   // ---------- 网络 20 ----------
   // 标题：*************故障计数（包含水平钻超时，凿超时，低电流，打孔深度超限）***********************
   // 注释：VisualChiseling No Sloping Hammer, added not  DB2500.DBX30.0  and #DrillHorizontal.StopDrill_Ack (in Network End) by WXY, 20220726
   // 含义：调用计数器实例 "Timer_DrilEndPos".TON（上升沿计数，当前值写入 CV）
   "Timer_DrilEndPos".TON(IN := (((((#HorDrillStep.S20 AND NOT (#HorDrillStep.S22)) OR ((#HorDrillStep.S22 AND NOT (#HorDrillStep.S25)) AND NOT ("DB2500 Visual Chiseling".VisualChiselingMode))) AND "DB1900_Communication_PC".Para.ProduceMode3) AND "DB720_KuKa_MainCtrl".StatusIn.do_DrilEnd_Pos) AND ("DB1900_Communication_PC".Recv.Current_2 < "DB1900_Communication_PC".Para.CurrentMinLimit)),
                          PT := T#2s);
   // 含义：条件 "Timer_DrilEndPos".Q 成立时，将 TRUE 传送到 "DB2500 Visual Chiseling".VChiselEndPos
   IF "Timer_DrilEndPos".Q THEN
       "DB2500 Visual Chiseling".VChiselEndPos := TRUE;
   END_IF;
   // 含义：条件 "Timer_DrilEndPos".Q 成立时，将 ("DB1042_Timer".HCLowTimeOutTimes + 1) 传送到 "DB1042_Timer".HCLowTimeOutTimes
   IF "Timer_DrilEndPos".Q THEN
       "DB1042_Timer".HCLowTimeOutTimes := ("DB1042_Timer".HCLowTimeOutTimes + 1);
   END_IF;
   // 含义：条件 ((((((#HorDrillStep.S20 AND NOT (#HorDrillStep.S22)) OR ((#HorDrillStep.S22 AND NOT (#HorDrillStep.S25)) AND NOT ("DB2500 Visual Chiseling".VisualChiselingMode))) AND "DB1900_Communication_PC".Para.ProduceMode3) AND ("DB1900_Communication_PC".Recv.Current_2 > "DB1900_Communication_PC".Para.CurrentMinLimit))) AND ("DB1900_Communication_PC".Recv.Current_2 < "DB1900_Communication_PC".Para.CurrentMaxLimit)) 成立时，将 0 传送到 "DB1042_Timer".HCLowTimeOutTimes
   IF ((((((#HorDrillStep.S20 AND NOT (#HorDrillStep.S22)) OR ((#HorDrillStep.S22 AND NOT (#HorDrillStep.S25)) AND NOT ("DB2500 Visual Chiseling".VisualChiselingMode))) AND "DB1900_Communication_PC".Para.ProduceMode3) AND ("DB1900_Communication_PC".Recv.Current_2 > "DB1900_Communication_PC".Para.CurrentMinLimit))) AND ("DB1900_Communication_PC".Recv.Current_2 < "DB1900_Communication_PC".Para.CurrentMaxLimit)) THEN
       "DB1042_Timer".HCLowTimeOutTimes := 0;
   END_IF;
   // 含义：条件 (((((#HorDrillStep.S20 AND NOT (#HorDrillStep.S22)) OR ((#HorDrillStep.S22 AND NOT (#HorDrillStep.S25)) AND NOT ("DB2500 Visual Chiseling".VisualChiselingMode))) AND "DB1900_Communication_PC".Para.ProduceMode3) AND "DB1042_Timer".HDrillEndTime.Q) OR ((((#HorDrillStep.S20 AND NOT (#HorDrillStep.S22)) OR ((#HorDrillStep.S22 AND NOT (#HorDrillStep.S25)) AND NOT ("DB2500 Visual Chiseling".VisualChiselingMode))) AND "DB1900_Communication_PC".Para.ProduceMode3) AND "DB1042_Timer".GougeTimeOut.Q) OR ((((#HorDrillStep.S20 AND NOT (#HorDrillStep.S22)) OR ((#HorDrillStep.S22 AND NOT (#HorDrillStep.S25)) AND NOT ("DB2500 Visual Chiseling".VisualChiselingMode))) AND "DB1900_Communication_PC".Para.ProduceMode3) AND "DB1042_Timer".CurrentLowTimeOut.Q) OR ((((#HorDrillStep.S20 AND NOT (#HorDrillStep.S22)) OR ((#HorDrillStep.S22 AND NOT (#HorDrillStep.S25)) AND NOT ("DB2500 Visual Chiseling".VisualChiselingMode))) AND "DB1900_Communication_PC".Para.ProduceMode3) AND "DB1042_Timer".CurrentHighTimeOut.Q) OR (((((#HorDrillStep.S20 AND NOT (#HorDrillStep.S22)) OR ((#HorDrillStep.S22 AND NOT (#HorDrillStep.S25)) AND NOT ("DB2500 Visual Chiseling".VisualChiselingMode))) AND "DB1900_Communication_PC".Para.ProduceMode3) AND ("DB1900_Communication_PC".Send.ScrLen >= "DB1900_Communication_PC".Para.DrillDepth))) OR ((((#HorDrillStep.S20 AND NOT (#HorDrillStep.S22)) OR ((#HorDrillStep.S22 AND NOT (#HorDrillStep.S25)) AND NOT ("DB2500 Visual Chiseling".VisualChiselingMode))) AND "DB1900_Communication_PC".Para.ProduceMode3) AND "DB2500 Visual Chiseling".VChiselEndPos)) AND NOT ("DB720_KuKa_MainCtrl".StatusIn.do_ChiselCylinderExt) 成立时，将 0.1 传送到 "DB1080_Component".Aux.Pressure
   IF (((((#HorDrillStep.S20 AND NOT (#HorDrillStep.S22)) OR ((#HorDrillStep.S22 AND NOT (#HorDrillStep.S25)) AND NOT ("DB2500 Visual Chiseling".VisualChiselingMode))) AND "DB1900_Communication_PC".Para.ProduceMode3) AND "DB1042_Timer".HDrillEndTime.Q) OR ((((#HorDrillStep.S20 AND NOT (#HorDrillStep.S22)) OR ((#HorDrillStep.S22 AND NOT (#HorDrillStep.S25)) AND NOT ("DB2500 Visual Chiseling".VisualChiselingMode))) AND "DB1900_Communication_PC".Para.ProduceMode3) AND "DB1042_Timer".GougeTimeOut.Q) OR ((((#HorDrillStep.S20 AND NOT (#HorDrillStep.S22)) OR ((#HorDrillStep.S22 AND NOT (#HorDrillStep.S25)) AND NOT ("DB2500 Visual Chiseling".VisualChiselingMode))) AND "DB1900_Communication_PC".Para.ProduceMode3) AND "DB1042_Timer".CurrentLowTimeOut.Q) OR ((((#HorDrillStep.S20 AND NOT (#HorDrillStep.S22)) OR ((#HorDrillStep.S22 AND NOT (#HorDrillStep.S25)) AND NOT ("DB2500 Visual Chiseling".VisualChiselingMode))) AND "DB1900_Communication_PC".Para.ProduceMode3) AND "DB1042_Timer".CurrentHighTimeOut.Q) OR (((((#HorDrillStep.S20 AND NOT (#HorDrillStep.S22)) OR ((#HorDrillStep.S22 AND NOT (#HorDrillStep.S25)) AND NOT ("DB2500 Visual Chiseling".VisualChiselingMode))) AND "DB1900_Communication_PC".Para.ProduceMode3) AND ("DB1900_Communication_PC".Send.ScrLen >= "DB1900_Communication_PC".Para.DrillDepth))) OR ((((#HorDrillStep.S20 AND NOT (#HorDrillStep.S22)) OR ((#HorDrillStep.S22 AND NOT (#HorDrillStep.S25)) AND NOT ("DB2500 Visual Chiseling".VisualChiselingMode))) AND "DB1900_Communication_PC".Para.ProduceMode3) AND "DB2500 Visual Chiseling".VChiselEndPos)) AND NOT ("DB720_KuKa_MainCtrl".StatusIn.do_ChiselCylinderExt) THEN
       "DB1080_Component".Aux.Pressure := 0.1;
   END_IF;
   // 含义：条件 (((((#HorDrillStep.S20 AND NOT (#HorDrillStep.S22)) OR ((#HorDrillStep.S22 AND NOT (#HorDrillStep.S25)) AND NOT ("DB2500 Visual Chiseling".VisualChiselingMode))) AND "DB1900_Communication_PC".Para.ProduceMode3) AND "DB1042_Timer".HDrillEndTime.Q) OR ((((#HorDrillStep.S20 AND NOT (#HorDrillStep.S22)) OR ((#HorDrillStep.S22 AND NOT (#HorDrillStep.S25)) AND NOT ("DB2500 Visual Chiseling".VisualChiselingMode))) AND "DB1900_Communication_PC".Para.ProduceMode3) AND "DB1042_Timer".GougeTimeOut.Q) OR ((((#HorDrillStep.S20 AND NOT (#HorDrillStep.S22)) OR ((#HorDrillStep.S22 AND NOT (#HorDrillStep.S25)) AND NOT ("DB2500 Visual Chiseling".VisualChiselingMode))) AND "DB1900_Communication_PC".Para.ProduceMode3) AND "DB1042_Timer".CurrentLowTimeOut.Q) OR ((((#HorDrillStep.S20 AND NOT (#HorDrillStep.S22)) OR ((#HorDrillStep.S22 AND NOT (#HorDrillStep.S25)) AND NOT ("DB2500 Visual Chiseling".VisualChiselingMode))) AND "DB1900_Communication_PC".Para.ProduceMode3) AND "DB1042_Timer".CurrentHighTimeOut.Q) OR (((((#HorDrillStep.S20 AND NOT (#HorDrillStep.S22)) OR ((#HorDrillStep.S22 AND NOT (#HorDrillStep.S25)) AND NOT ("DB2500 Visual Chiseling".VisualChiselingMode))) AND "DB1900_Communication_PC".Para.ProduceMode3) AND ("DB1900_Communication_PC".Send.ScrLen >= "DB1900_Communication_PC".Para.DrillDepth))) OR ((((#HorDrillStep.S20 AND NOT (#HorDrillStep.S22)) OR ((#HorDrillStep.S22 AND NOT (#HorDrillStep.S25)) AND NOT ("DB2500 Visual Chiseling".VisualChiselingMode))) AND "DB1900_Communication_PC".Para.ProduceMode3) AND "DB2500 Visual Chiseling".VChiselEndPos)) AND NOT ("DB720_KuKa_MainCtrl".CmdOut.di_ChiselRobotRet) 成立时，将 TRUE 传送到 "DB1081_ValveCall".ST01.Z02.RetAuto
   IF (((((#HorDrillStep.S20 AND NOT (#HorDrillStep.S22)) OR ((#HorDrillStep.S22 AND NOT (#HorDrillStep.S25)) AND NOT ("DB2500 Visual Chiseling".VisualChiselingMode))) AND "DB1900_Communication_PC".Para.ProduceMode3) AND "DB1042_Timer".HDrillEndTime.Q) OR ((((#HorDrillStep.S20 AND NOT (#HorDrillStep.S22)) OR ((#HorDrillStep.S22 AND NOT (#HorDrillStep.S25)) AND NOT ("DB2500 Visual Chiseling".VisualChiselingMode))) AND "DB1900_Communication_PC".Para.ProduceMode3) AND "DB1042_Timer".GougeTimeOut.Q) OR ((((#HorDrillStep.S20 AND NOT (#HorDrillStep.S22)) OR ((#HorDrillStep.S22 AND NOT (#HorDrillStep.S25)) AND NOT ("DB2500 Visual Chiseling".VisualChiselingMode))) AND "DB1900_Communication_PC".Para.ProduceMode3) AND "DB1042_Timer".CurrentLowTimeOut.Q) OR ((((#HorDrillStep.S20 AND NOT (#HorDrillStep.S22)) OR ((#HorDrillStep.S22 AND NOT (#HorDrillStep.S25)) AND NOT ("DB2500 Visual Chiseling".VisualChiselingMode))) AND "DB1900_Communication_PC".Para.ProduceMode3) AND "DB1042_Timer".CurrentHighTimeOut.Q) OR (((((#HorDrillStep.S20 AND NOT (#HorDrillStep.S22)) OR ((#HorDrillStep.S22 AND NOT (#HorDrillStep.S25)) AND NOT ("DB2500 Visual Chiseling".VisualChiselingMode))) AND "DB1900_Communication_PC".Para.ProduceMode3) AND ("DB1900_Communication_PC".Send.ScrLen >= "DB1900_Communication_PC".Para.DrillDepth))) OR ((((#HorDrillStep.S20 AND NOT (#HorDrillStep.S22)) OR ((#HorDrillStep.S22 AND NOT (#HorDrillStep.S25)) AND NOT ("DB2500 Visual Chiseling".VisualChiselingMode))) AND "DB1900_Communication_PC".Para.ProduceMode3) AND "DB2500 Visual Chiseling".VChiselEndPos)) AND NOT ("DB720_KuKa_MainCtrl".CmdOut.di_ChiselRobotRet) THEN
       "DB1081_ValveCall".ST01.Z02.RetAuto := TRUE;
   END_IF;
   // 含义：条件 (((((#HorDrillStep.S20 AND NOT (#HorDrillStep.S22)) OR ((#HorDrillStep.S22 AND NOT (#HorDrillStep.S25)) AND NOT ("DB2500 Visual Chiseling".VisualChiselingMode))) AND "DB1900_Communication_PC".Para.ProduceMode3) AND "DB1042_Timer".HDrillEndTime.Q) OR ((((#HorDrillStep.S20 AND NOT (#HorDrillStep.S22)) OR ((#HorDrillStep.S22 AND NOT (#HorDrillStep.S25)) AND NOT ("DB2500 Visual Chiseling".VisualChiselingMode))) AND "DB1900_Communication_PC".Para.ProduceMode3) AND "DB1042_Timer".GougeTimeOut.Q) OR ((((#HorDrillStep.S20 AND NOT (#HorDrillStep.S22)) OR ((#HorDrillStep.S22 AND NOT (#HorDrillStep.S25)) AND NOT ("DB2500 Visual Chiseling".VisualChiselingMode))) AND "DB1900_Communication_PC".Para.ProduceMode3) AND "DB1042_Timer".CurrentLowTimeOut.Q) OR ((((#HorDrillStep.S20 AND NOT (#HorDrillStep.S22)) OR ((#HorDrillStep.S22 AND NOT (#HorDrillStep.S25)) AND NOT ("DB2500 Visual Chiseling".VisualChiselingMode))) AND "DB1900_Communication_PC".Para.ProduceMode3) AND "DB1042_Timer".CurrentHighTimeOut.Q) OR (((((#HorDrillStep.S20 AND NOT (#HorDrillStep.S22)) OR ((#HorDrillStep.S22 AND NOT (#HorDrillStep.S25)) AND NOT ("DB2500 Visual Chiseling".VisualChiselingMode))) AND "DB1900_Communication_PC".Para.ProduceMode3) AND ("DB1900_Communication_PC".Send.ScrLen >= "DB1900_Communication_PC".Para.DrillDepth))) OR ((((#HorDrillStep.S20 AND NOT (#HorDrillStep.S22)) OR ((#HorDrillStep.S22 AND NOT (#HorDrillStep.S25)) AND NOT ("DB2500 Visual Chiseling".VisualChiselingMode))) AND "DB1900_Communication_PC".Para.ProduceMode3) AND "DB2500 Visual Chiseling".VChiselEndPos)) AND "DB720_KuKa_MainCtrl".StatusIn.do_ChiselCylinderExt 成立时，将 FALSE 传送到 "DB1081_ValveCall".ST01.Z02.RetAuto
   IF (((((#HorDrillStep.S20 AND NOT (#HorDrillStep.S22)) OR ((#HorDrillStep.S22 AND NOT (#HorDrillStep.S25)) AND NOT ("DB2500 Visual Chiseling".VisualChiselingMode))) AND "DB1900_Communication_PC".Para.ProduceMode3) AND "DB1042_Timer".HDrillEndTime.Q) OR ((((#HorDrillStep.S20 AND NOT (#HorDrillStep.S22)) OR ((#HorDrillStep.S22 AND NOT (#HorDrillStep.S25)) AND NOT ("DB2500 Visual Chiseling".VisualChiselingMode))) AND "DB1900_Communication_PC".Para.ProduceMode3) AND "DB1042_Timer".GougeTimeOut.Q) OR ((((#HorDrillStep.S20 AND NOT (#HorDrillStep.S22)) OR ((#HorDrillStep.S22 AND NOT (#HorDrillStep.S25)) AND NOT ("DB2500 Visual Chiseling".VisualChiselingMode))) AND "DB1900_Communication_PC".Para.ProduceMode3) AND "DB1042_Timer".CurrentLowTimeOut.Q) OR ((((#HorDrillStep.S20 AND NOT (#HorDrillStep.S22)) OR ((#HorDrillStep.S22 AND NOT (#HorDrillStep.S25)) AND NOT ("DB2500 Visual Chiseling".VisualChiselingMode))) AND "DB1900_Communication_PC".Para.ProduceMode3) AND "DB1042_Timer".CurrentHighTimeOut.Q) OR (((((#HorDrillStep.S20 AND NOT (#HorDrillStep.S22)) OR ((#HorDrillStep.S22 AND NOT (#HorDrillStep.S25)) AND NOT ("DB2500 Visual Chiseling".VisualChiselingMode))) AND "DB1900_Communication_PC".Para.ProduceMode3) AND ("DB1900_Communication_PC".Send.ScrLen >= "DB1900_Communication_PC".Para.DrillDepth))) OR ((((#HorDrillStep.S20 AND NOT (#HorDrillStep.S22)) OR ((#HorDrillStep.S22 AND NOT (#HorDrillStep.S25)) AND NOT ("DB2500 Visual Chiseling".VisualChiselingMode))) AND "DB1900_Communication_PC".Para.ProduceMode3) AND "DB2500 Visual Chiseling".VChiselEndPos)) AND "DB720_KuKa_MainCtrl".StatusIn.do_ChiselCylinderExt THEN
       "DB1081_ValveCall".ST01.Z02.RetAuto := FALSE;
   END_IF;
   // 含义：条件 (((((#HorDrillStep.S20 AND NOT (#HorDrillStep.S22)) OR ((#HorDrillStep.S22 AND NOT (#HorDrillStep.S25)) AND NOT ("DB2500 Visual Chiseling".VisualChiselingMode))) AND "DB1900_Communication_PC".Para.ProduceMode3) AND "DB1042_Timer".HDrillEndTime.Q) OR ((((#HorDrillStep.S20 AND NOT (#HorDrillStep.S22)) OR ((#HorDrillStep.S22 AND NOT (#HorDrillStep.S25)) AND NOT ("DB2500 Visual Chiseling".VisualChiselingMode))) AND "DB1900_Communication_PC".Para.ProduceMode3) AND "DB1042_Timer".GougeTimeOut.Q) OR ((((#HorDrillStep.S20 AND NOT (#HorDrillStep.S22)) OR ((#HorDrillStep.S22 AND NOT (#HorDrillStep.S25)) AND NOT ("DB2500 Visual Chiseling".VisualChiselingMode))) AND "DB1900_Communication_PC".Para.ProduceMode3) AND "DB1042_Timer".CurrentLowTimeOut.Q) OR ((((#HorDrillStep.S20 AND NOT (#HorDrillStep.S22)) OR ((#HorDrillStep.S22 AND NOT (#HorDrillStep.S25)) AND NOT ("DB2500 Visual Chiseling".VisualChiselingMode))) AND "DB1900_Communication_PC".Para.ProduceMode3) AND "DB1042_Timer".CurrentHighTimeOut.Q) OR (((((#HorDrillStep.S20 AND NOT (#HorDrillStep.S22)) OR ((#HorDrillStep.S22 AND NOT (#HorDrillStep.S25)) AND NOT ("DB2500 Visual Chiseling".VisualChiselingMode))) AND "DB1900_Communication_PC".Para.ProduceMode3) AND ("DB1900_Communication_PC".Send.ScrLen >= "DB1900_Communication_PC".Para.DrillDepth))) OR ((((#HorDrillStep.S20 AND NOT (#HorDrillStep.S22)) OR ((#HorDrillStep.S22 AND NOT (#HorDrillStep.S25)) AND NOT ("DB2500 Visual Chiseling".VisualChiselingMode))) AND "DB1900_Communication_PC".Para.ProduceMode3) AND "DB2500 Visual Chiseling".VChiselEndPos)) AND "DB720_KuKa_MainCtrl".StatusIn.do_ReqStopDril 成立时，将 FALSE 传送到 "DB720_KuKa_MainCtrl".CmdOut.di_ChiselCylinderRet
   IF (((((#HorDrillStep.S20 AND NOT (#HorDrillStep.S22)) OR ((#HorDrillStep.S22 AND NOT (#HorDrillStep.S25)) AND NOT ("DB2500 Visual Chiseling".VisualChiselingMode))) AND "DB1900_Communication_PC".Para.ProduceMode3) AND "DB1042_Timer".HDrillEndTime.Q) OR ((((#HorDrillStep.S20 AND NOT (#HorDrillStep.S22)) OR ((#HorDrillStep.S22 AND NOT (#HorDrillStep.S25)) AND NOT ("DB2500 Visual Chiseling".VisualChiselingMode))) AND "DB1900_Communication_PC".Para.ProduceMode3) AND "DB1042_Timer".GougeTimeOut.Q) OR ((((#HorDrillStep.S20 AND NOT (#HorDrillStep.S22)) OR ((#HorDrillStep.S22 AND NOT (#HorDrillStep.S25)) AND NOT ("DB2500 Visual Chiseling".VisualChiselingMode))) AND "DB1900_Communication_PC".Para.ProduceMode3) AND "DB1042_Timer".CurrentLowTimeOut.Q) OR ((((#HorDrillStep.S20 AND NOT (#HorDrillStep.S22)) OR ((#HorDrillStep.S22 AND NOT (#HorDrillStep.S25)) AND NOT ("DB2500 Visual Chiseling".VisualChiselingMode))) AND "DB1900_Communication_PC".Para.ProduceMode3) AND "DB1042_Timer".CurrentHighTimeOut.Q) OR (((((#HorDrillStep.S20 AND NOT (#HorDrillStep.S22)) OR ((#HorDrillStep.S22 AND NOT (#HorDrillStep.S25)) AND NOT ("DB2500 Visual Chiseling".VisualChiselingMode))) AND "DB1900_Communication_PC".Para.ProduceMode3) AND ("DB1900_Communication_PC".Send.ScrLen >= "DB1900_Communication_PC".Para.DrillDepth))) OR ((((#HorDrillStep.S20 AND NOT (#HorDrillStep.S22)) OR ((#HorDrillStep.S22 AND NOT (#HorDrillStep.S25)) AND NOT ("DB2500 Visual Chiseling".VisualChiselingMode))) AND "DB1900_Communication_PC".Para.ProduceMode3) AND "DB2500 Visual Chiseling".VChiselEndPos)) AND "DB720_KuKa_MainCtrl".StatusIn.do_ReqStopDril THEN
       "DB720_KuKa_MainCtrl".CmdOut.di_ChiselCylinderRet := FALSE;
   END_IF;
   // 含义：条件 (((((#HorDrillStep.S20 AND NOT (#HorDrillStep.S22)) OR ((#HorDrillStep.S22 AND NOT (#HorDrillStep.S25)) AND NOT ("DB2500 Visual Chiseling".VisualChiselingMode))) AND "DB1900_Communication_PC".Para.ProduceMode3) AND "DB1042_Timer".HDrillEndTime.Q) OR ((((#HorDrillStep.S20 AND NOT (#HorDrillStep.S22)) OR ((#HorDrillStep.S22 AND NOT (#HorDrillStep.S25)) AND NOT ("DB2500 Visual Chiseling".VisualChiselingMode))) AND "DB1900_Communication_PC".Para.ProduceMode3) AND "DB1042_Timer".GougeTimeOut.Q) OR ((((#HorDrillStep.S20 AND NOT (#HorDrillStep.S22)) OR ((#HorDrillStep.S22 AND NOT (#HorDrillStep.S25)) AND NOT ("DB2500 Visual Chiseling".VisualChiselingMode))) AND "DB1900_Communication_PC".Para.ProduceMode3) AND "DB1042_Timer".CurrentLowTimeOut.Q) OR ((((#HorDrillStep.S20 AND NOT (#HorDrillStep.S22)) OR ((#HorDrillStep.S22 AND NOT (#HorDrillStep.S25)) AND NOT ("DB2500 Visual Chiseling".VisualChiselingMode))) AND "DB1900_Communication_PC".Para.ProduceMode3) AND "DB1042_Timer".CurrentHighTimeOut.Q) OR (((((#HorDrillStep.S20 AND NOT (#HorDrillStep.S22)) OR ((#HorDrillStep.S22 AND NOT (#HorDrillStep.S25)) AND NOT ("DB2500 Visual Chiseling".VisualChiselingMode))) AND "DB1900_Communication_PC".Para.ProduceMode3) AND ("DB1900_Communication_PC".Send.ScrLen >= "DB1900_Communication_PC".Para.DrillDepth))) OR ((((#HorDrillStep.S20 AND NOT (#HorDrillStep.S22)) OR ((#HorDrillStep.S22 AND NOT (#HorDrillStep.S25)) AND NOT ("DB2500 Visual Chiseling".VisualChiselingMode))) AND "DB1900_Communication_PC".Para.ProduceMode3) AND "DB2500 Visual Chiseling".VChiselEndPos)) AND "DB720_KuKa_MainCtrl".StatusIn.do_ReqStopDril 成立时，将 FALSE 传送到 "DB720_KuKa_MainCtrl".CmdOut.di_ChiselRobotRet
   IF (((((#HorDrillStep.S20 AND NOT (#HorDrillStep.S22)) OR ((#HorDrillStep.S22 AND NOT (#HorDrillStep.S25)) AND NOT ("DB2500 Visual Chiseling".VisualChiselingMode))) AND "DB1900_Communication_PC".Para.ProduceMode3) AND "DB1042_Timer".HDrillEndTime.Q) OR ((((#HorDrillStep.S20 AND NOT (#HorDrillStep.S22)) OR ((#HorDrillStep.S22 AND NOT (#HorDrillStep.S25)) AND NOT ("DB2500 Visual Chiseling".VisualChiselingMode))) AND "DB1900_Communication_PC".Para.ProduceMode3) AND "DB1042_Timer".GougeTimeOut.Q) OR ((((#HorDrillStep.S20 AND NOT (#HorDrillStep.S22)) OR ((#HorDrillStep.S22 AND NOT (#HorDrillStep.S25)) AND NOT ("DB2500 Visual Chiseling".VisualChiselingMode))) AND "DB1900_Communication_PC".Para.ProduceMode3) AND "DB1042_Timer".CurrentLowTimeOut.Q) OR ((((#HorDrillStep.S20 AND NOT (#HorDrillStep.S22)) OR ((#HorDrillStep.S22 AND NOT (#HorDrillStep.S25)) AND NOT ("DB2500 Visual Chiseling".VisualChiselingMode))) AND "DB1900_Communication_PC".Para.ProduceMode3) AND "DB1042_Timer".CurrentHighTimeOut.Q) OR (((((#HorDrillStep.S20 AND NOT (#HorDrillStep.S22)) OR ((#HorDrillStep.S22 AND NOT (#HorDrillStep.S25)) AND NOT ("DB2500 Visual Chiseling".VisualChiselingMode))) AND "DB1900_Communication_PC".Para.ProduceMode3) AND ("DB1900_Communication_PC".Send.ScrLen >= "DB1900_Communication_PC".Para.DrillDepth))) OR ((((#HorDrillStep.S20 AND NOT (#HorDrillStep.S22)) OR ((#HorDrillStep.S22 AND NOT (#HorDrillStep.S25)) AND NOT ("DB2500 Visual Chiseling".VisualChiselingMode))) AND "DB1900_Communication_PC".Para.ProduceMode3) AND "DB2500 Visual Chiseling".VChiselEndPos)) AND "DB720_KuKa_MainCtrl".StatusIn.do_ReqStopDril THEN
       "DB720_KuKa_MainCtrl".CmdOut.di_ChiselRobotRet := FALSE;
   END_IF;
   // 含义：条件 (((((((#HorDrillStep.S20 AND NOT (#HorDrillStep.S22)) OR ((#HorDrillStep.S22 AND NOT (#HorDrillStep.S25)) AND NOT ("DB2500 Visual Chiseling".VisualChiselingMode))) AND "DB1900_Communication_PC".Para.ProduceMode3) AND "DB1042_Timer".HDrillEndTime.Q) OR ((((#HorDrillStep.S20 AND NOT (#HorDrillStep.S22)) OR ((#HorDrillStep.S22 AND NOT (#HorDrillStep.S25)) AND NOT ("DB2500 Visual Chiseling".VisualChiselingMode))) AND "DB1900_Communication_PC".Para.ProduceMode3) AND "DB1042_Timer".GougeTimeOut.Q) OR ((((#HorDrillStep.S20 AND NOT (#HorDrillStep.S22)) OR ((#HorDrillStep.S22 AND NOT (#HorDrillStep.S25)) AND NOT ("DB2500 Visual Chiseling".VisualChiselingMode))) AND "DB1900_Communication_PC".Para.ProduceMode3) AND "DB1042_Timer".CurrentLowTimeOut.Q) OR ((((#HorDrillStep.S20 AND NOT (#HorDrillStep.S22)) OR ((#HorDrillStep.S22 AND NOT (#HorDrillStep.S25)) AND NOT ("DB2500 Visual Chiseling".VisualChiselingMode))) AND "DB1900_Communication_PC".Para.ProduceMode3) AND "DB1042_Timer".CurrentHighTimeOut.Q) OR (((((#HorDrillStep.S20 AND NOT (#HorDrillStep.S22)) OR ((#HorDrillStep.S22 AND NOT (#HorDrillStep.S25)) AND NOT ("DB2500 Visual Chiseling".VisualChiselingMode))) AND "DB1900_Communication_PC".Para.ProduceMode3) AND ("DB1900_Communication_PC".Send.ScrLen >= "DB1900_Communication_PC".Para.DrillDepth))) OR ((((#HorDrillStep.S20 AND NOT (#HorDrillStep.S22)) OR ((#HorDrillStep.S22 AND NOT (#HorDrillStep.S25)) AND NOT ("DB2500 Visual Chiseling".VisualChiselingMode))) AND "DB1900_Communication_PC".Para.ProduceMode3) AND "DB2500 Visual Chiseling".VChiselEndPos)) AND "IZ02RetPos") AND ("DB1080_Component".ClinyderPos.Ctrl_Out.Cur_Val_Out >= 92.5)) 成立时，将 TRUE 传送到 "DB720_KuKa_MainCtrl".CmdOut.di_ChiselRobotRet
   IF (((((((#HorDrillStep.S20 AND NOT (#HorDrillStep.S22)) OR ((#HorDrillStep.S22 AND NOT (#HorDrillStep.S25)) AND NOT ("DB2500 Visual Chiseling".VisualChiselingMode))) AND "DB1900_Communication_PC".Para.ProduceMode3) AND "DB1042_Timer".HDrillEndTime.Q) OR ((((#HorDrillStep.S20 AND NOT (#HorDrillStep.S22)) OR ((#HorDrillStep.S22 AND NOT (#HorDrillStep.S25)) AND NOT ("DB2500 Visual Chiseling".VisualChiselingMode))) AND "DB1900_Communication_PC".Para.ProduceMode3) AND "DB1042_Timer".GougeTimeOut.Q) OR ((((#HorDrillStep.S20 AND NOT (#HorDrillStep.S22)) OR ((#HorDrillStep.S22 AND NOT (#HorDrillStep.S25)) AND NOT ("DB2500 Visual Chiseling".VisualChiselingMode))) AND "DB1900_Communication_PC".Para.ProduceMode3) AND "DB1042_Timer".CurrentLowTimeOut.Q) OR ((((#HorDrillStep.S20 AND NOT (#HorDrillStep.S22)) OR ((#HorDrillStep.S22 AND NOT (#HorDrillStep.S25)) AND NOT ("DB2500 Visual Chiseling".VisualChiselingMode))) AND "DB1900_Communication_PC".Para.ProduceMode3) AND "DB1042_Timer".CurrentHighTimeOut.Q) OR (((((#HorDrillStep.S20 AND NOT (#HorDrillStep.S22)) OR ((#HorDrillStep.S22 AND NOT (#HorDrillStep.S25)) AND NOT ("DB2500 Visual Chiseling".VisualChiselingMode))) AND "DB1900_Communication_PC".Para.ProduceMode3) AND ("DB1900_Communication_PC".Send.ScrLen >= "DB1900_Communication_PC".Para.DrillDepth))) OR ((((#HorDrillStep.S20 AND NOT (#HorDrillStep.S22)) OR ((#HorDrillStep.S22 AND NOT (#HorDrillStep.S25)) AND NOT ("DB2500 Visual Chiseling".VisualChiselingMode))) AND "DB1900_Communication_PC".Para.ProduceMode3) AND "DB2500 Visual Chiseling".VChiselEndPos)) AND "IZ02RetPos") AND ("DB1080_Component".ClinyderPos.Ctrl_Out.Cur_Val_Out >= 92.5)) THEN
       "DB720_KuKa_MainCtrl".CmdOut.di_ChiselRobotRet := TRUE;
   END_IF;
   // 含义：条件 (((((((#HorDrillStep.S20 AND NOT (#HorDrillStep.S22)) OR ((#HorDrillStep.S22 AND NOT (#HorDrillStep.S25)) AND NOT ("DB2500 Visual Chiseling".VisualChiselingMode))) AND "DB1900_Communication_PC".Para.ProduceMode3) AND "DB1042_Timer".HDrillEndTime.Q) OR ((((#HorDrillStep.S20 AND NOT (#HorDrillStep.S22)) OR ((#HorDrillStep.S22 AND NOT (#HorDrillStep.S25)) AND NOT ("DB2500 Visual Chiseling".VisualChiselingMode))) AND "DB1900_Communication_PC".Para.ProduceMode3) AND "DB1042_Timer".GougeTimeOut.Q) OR ((((#HorDrillStep.S20 AND NOT (#HorDrillStep.S22)) OR ((#HorDrillStep.S22 AND NOT (#HorDrillStep.S25)) AND NOT ("DB2500 Visual Chiseling".VisualChiselingMode))) AND "DB1900_Communication_PC".Para.ProduceMode3) AND "DB1042_Timer".CurrentLowTimeOut.Q) OR ((((#HorDrillStep.S20 AND NOT (#HorDrillStep.S22)) OR ((#HorDrillStep.S22 AND NOT (#HorDrillStep.S25)) AND NOT ("DB2500 Visual Chiseling".VisualChiselingMode))) AND "DB1900_Communication_PC".Para.ProduceMode3) AND "DB1042_Timer".CurrentHighTimeOut.Q) OR (((((#HorDrillStep.S20 AND NOT (#HorDrillStep.S22)) OR ((#HorDrillStep.S22 AND NOT (#HorDrillStep.S25)) AND NOT ("DB2500 Visual Chiseling".VisualChiselingMode))) AND "DB1900_Communication_PC".Para.ProduceMode3) AND ("DB1900_Communication_PC".Send.ScrLen >= "DB1900_Communication_PC".Para.DrillDepth))) OR ((((#HorDrillStep.S20 AND NOT (#HorDrillStep.S22)) OR ((#HorDrillStep.S22 AND NOT (#HorDrillStep.S25)) AND NOT ("DB2500 Visual Chiseling".VisualChiselingMode))) AND "DB1900_Communication_PC".Para.ProduceMode3) AND "DB2500 Visual Chiseling".VChiselEndPos)) AND "IZ02RetPos") AND ("DB1080_Component".ClinyderPos.Ctrl_Out.Cur_Val_Out >= 92.5)) 成立时，将 TRUE 传送到 "DB720_KuKa_MainCtrl".CmdOut.di_ChiselCylinderRet
   IF (((((((#HorDrillStep.S20 AND NOT (#HorDrillStep.S22)) OR ((#HorDrillStep.S22 AND NOT (#HorDrillStep.S25)) AND NOT ("DB2500 Visual Chiseling".VisualChiselingMode))) AND "DB1900_Communication_PC".Para.ProduceMode3) AND "DB1042_Timer".HDrillEndTime.Q) OR ((((#HorDrillStep.S20 AND NOT (#HorDrillStep.S22)) OR ((#HorDrillStep.S22 AND NOT (#HorDrillStep.S25)) AND NOT ("DB2500 Visual Chiseling".VisualChiselingMode))) AND "DB1900_Communication_PC".Para.ProduceMode3) AND "DB1042_Timer".GougeTimeOut.Q) OR ((((#HorDrillStep.S20 AND NOT (#HorDrillStep.S22)) OR ((#HorDrillStep.S22 AND NOT (#HorDrillStep.S25)) AND NOT ("DB2500 Visual Chiseling".VisualChiselingMode))) AND "DB1900_Communication_PC".Para.ProduceMode3) AND "DB1042_Timer".CurrentLowTimeOut.Q) OR ((((#HorDrillStep.S20 AND NOT (#HorDrillStep.S22)) OR ((#HorDrillStep.S22 AND NOT (#HorDrillStep.S25)) AND NOT ("DB2500 Visual Chiseling".VisualChiselingMode))) AND "DB1900_Communication_PC".Para.ProduceMode3) AND "DB1042_Timer".CurrentHighTimeOut.Q) OR (((((#HorDrillStep.S20 AND NOT (#HorDrillStep.S22)) OR ((#HorDrillStep.S22 AND NOT (#HorDrillStep.S25)) AND NOT ("DB2500 Visual Chiseling".VisualChiselingMode))) AND "DB1900_Communication_PC".Para.ProduceMode3) AND ("DB1900_Communication_PC".Send.ScrLen >= "DB1900_Communication_PC".Para.DrillDepth))) OR ((((#HorDrillStep.S20 AND NOT (#HorDrillStep.S22)) OR ((#HorDrillStep.S22 AND NOT (#HorDrillStep.S25)) AND NOT ("DB2500 Visual Chiseling".VisualChiselingMode))) AND "DB1900_Communication_PC".Para.ProduceMode3) AND "DB2500 Visual Chiseling".VChiselEndPos)) AND "IZ02RetPos") AND ("DB1080_Component".ClinyderPos.Ctrl_Out.Cur_Val_Out >= 92.5)) THEN
       "DB720_KuKa_MainCtrl".CmdOut.di_ChiselCylinderRet := TRUE;
   END_IF;
   // 含义：调用计数器实例 "Timer_CylinderBack_Hor".TON（上升沿计数，当前值写入 CV）
   "Timer_CylinderBack_Hor".TON(IN := (((((#HorDrillStep.S20 AND NOT (#HorDrillStep.S22)) OR ((#HorDrillStep.S22 AND NOT (#HorDrillStep.S25)) AND NOT ("DB2500 Visual Chiseling".VisualChiselingMode))) AND "DB1900_Communication_PC".Para.ProduceMode3) AND "DB1042_Timer".HDrillEndTime.Q) OR ((((#HorDrillStep.S20 AND NOT (#HorDrillStep.S22)) OR ((#HorDrillStep.S22 AND NOT (#HorDrillStep.S25)) AND NOT ("DB2500 Visual Chiseling".VisualChiselingMode))) AND "DB1900_Communication_PC".Para.ProduceMode3) AND "DB1042_Timer".GougeTimeOut.Q) OR ((((#HorDrillStep.S20 AND NOT (#HorDrillStep.S22)) OR ((#HorDrillStep.S22 AND NOT (#HorDrillStep.S25)) AND NOT ("DB2500 Visual Chiseling".VisualChiselingMode))) AND "DB1900_Communication_PC".Para.ProduceMode3) AND "DB1042_Timer".CurrentLowTimeOut.Q) OR ((((#HorDrillStep.S20 AND NOT (#HorDrillStep.S22)) OR ((#HorDrillStep.S22 AND NOT (#HorDrillStep.S25)) AND NOT ("DB2500 Visual Chiseling".VisualChiselingMode))) AND "DB1900_Communication_PC".Para.ProduceMode3) AND "DB1042_Timer".CurrentHighTimeOut.Q) OR (((((#HorDrillStep.S20 AND NOT (#HorDrillStep.S22)) OR ((#HorDrillStep.S22 AND NOT (#HorDrillStep.S25)) AND NOT ("DB2500 Visual Chiseling".VisualChiselingMode))) AND "DB1900_Communication_PC".Para.ProduceMode3) AND ("DB1900_Communication_PC".Send.ScrLen >= "DB1900_Communication_PC".Para.DrillDepth))) OR ((((#HorDrillStep.S20 AND NOT (#HorDrillStep.S22)) OR ((#HorDrillStep.S22 AND NOT (#HorDrillStep.S25)) AND NOT ("DB2500 Visual Chiseling".VisualChiselingMode))) AND "DB1900_Communication_PC".Para.ProduceMode3) AND "DB2500 Visual Chiseling".VChiselEndPos)) AND NOT ("IZ02RetPos"),
                                PT := t#3s);
   // 含义：条件 "Timer_CylinderBack_Hor".Q 成立时，将 TRUE 传送到 "DB720_KuKa_MainCtrl".CmdOut.di_ChiselRobotRet
   IF "Timer_CylinderBack_Hor".Q THEN
       "DB720_KuKa_MainCtrl".CmdOut.di_ChiselRobotRet := TRUE;
   END_IF;
   // 含义：调用计数器实例 "Timer_RobotPry_Hor".TON（上升沿计数，当前值写入 CV）
   "Timer_RobotPry_Hor".TON(IN := ((((((#HorDrillStep.S20 AND NOT (#HorDrillStep.S22)) OR ((#HorDrillStep.S22 AND NOT (#HorDrillStep.S25)) AND NOT ("DB2500 Visual Chiseling".VisualChiselingMode))) AND "DB1900_Communication_PC".Para.ProduceMode3) AND "DB1042_Timer".HDrillEndTime.Q) OR ((((#HorDrillStep.S20 AND NOT (#HorDrillStep.S22)) OR ((#HorDrillStep.S22 AND NOT (#HorDrillStep.S25)) AND NOT ("DB2500 Visual Chiseling".VisualChiselingMode))) AND "DB1900_Communication_PC".Para.ProduceMode3) AND "DB1042_Timer".GougeTimeOut.Q) OR ((((#HorDrillStep.S20 AND NOT (#HorDrillStep.S22)) OR ((#HorDrillStep.S22 AND NOT (#HorDrillStep.S25)) AND NOT ("DB2500 Visual Chiseling".VisualChiselingMode))) AND "DB1900_Communication_PC".Para.ProduceMode3) AND "DB1042_Timer".CurrentLowTimeOut.Q) OR ((((#HorDrillStep.S20 AND NOT (#HorDrillStep.S22)) OR ((#HorDrillStep.S22 AND NOT (#HorDrillStep.S25)) AND NOT ("DB2500 Visual Chiseling".VisualChiselingMode))) AND "DB1900_Communication_PC".Para.ProduceMode3) AND "DB1042_Timer".CurrentHighTimeOut.Q) OR (((((#HorDrillStep.S20 AND NOT (#HorDrillStep.S22)) OR ((#HorDrillStep.S22 AND NOT (#HorDrillStep.S25)) AND NOT ("DB2500 Visual Chiseling".VisualChiselingMode))) AND "DB1900_Communication_PC".Para.ProduceMode3) AND ("DB1900_Communication_PC".Send.ScrLen >= "DB1900_Communication_PC".Para.DrillDepth))) OR ((((#HorDrillStep.S20 AND NOT (#HorDrillStep.S22)) OR ((#HorDrillStep.S22 AND NOT (#HorDrillStep.S25)) AND NOT ("DB2500 Visual Chiseling".VisualChiselingMode))) AND "DB1900_Communication_PC".Para.ProduceMode3) AND "DB2500 Visual Chiseling".VChiselEndPos)) AND NOT ("IZ02RetPos")) AND "DB720_KuKa_MainCtrl".StatusIn.do_RobotPry_End,
                            PT := t#3s);
   // 含义：条件 "Timer_RobotPry_Hor".Q 成立时，将 FALSE 传送到 "DB720_KuKa_MainCtrl".CmdOut.di_ChiselCylinderRet
   IF "Timer_RobotPry_Hor".Q THEN
       "DB720_KuKa_MainCtrl".CmdOut.di_ChiselCylinderRet := FALSE;
   END_IF;
   // 含义：条件 "Timer_RobotPry_Hor".Q 成立时，将 FALSE 传送到 "DB720_KuKa_MainCtrl".CmdOut.di_ChiselRobotRet
   IF "Timer_RobotPry_Hor".Q THEN
       "DB720_KuKa_MainCtrl".CmdOut.di_ChiselRobotRet := FALSE;
   END_IF;
   // 含义：条件 "Timer_RobotPry_Hor".Q 成立时，将 TRUE 传送到 #HorDrillStep.ErrEnd
   IF "Timer_RobotPry_Hor".Q THEN
       #HorDrillStep.ErrEnd := TRUE;
   END_IF;
   // 含义：条件 "Timer_RobotPry_Hor".Q 成立时，将 TRUE 传送到 "DB1148_PromptBeeper".Public.HorChiselStuckErr
   IF "Timer_RobotPry_Hor".Q THEN
       "DB1148_PromptBeeper".Public.HorChiselStuckErr := TRUE;
   END_IF;
   // 含义：条件 "Timer_RobotPry_Hor".Q 成立时，将 FALSE 传送到 "DB1081_ValveCall".ST01.Z02.RetAuto
   IF "Timer_RobotPry_Hor".Q THEN
       "DB1081_ValveCall".ST01.Z02.RetAuto := FALSE;
   END_IF;
   // 含义：条件 "Timer_RobotPry_Hor".Q 成立时，将 TRUE 传送到 "DB1081_ValveCall".ST01.Z01.ExtAuto
   IF "Timer_RobotPry_Hor".Q THEN
       "DB1081_ValveCall".ST01.Z01.ExtAuto := TRUE;
   END_IF;
   // 含义：条件 "Timer_RobotPry_Hor".Q 成立时，将 FALSE 传送到 "DB1081_ValveCall".ST01.Z01.RetAuto
   IF "Timer_RobotPry_Hor".Q THEN
       "DB1081_ValveCall".ST01.Z01.RetAuto := FALSE;
   END_IF;
   // 含义：条件 "Timer_RobotPry_Hor".Q 成立时，将 0.5 传送到 "DB1080_Component".Aux.Pressure
   IF "Timer_RobotPry_Hor".Q THEN
       "DB1080_Component".Aux.Pressure := 0.5;
   END_IF;
   // 含义：将 ((((#HorDrillStep.S20 AND NOT (#HorDrillStep.S22)) OR ((#HorDrillStep.S22 AND NOT (#HorDrillStep.S25)) AND NOT ("DB2500 Visual Chiseling".VisualChiselingMode))) AND "DB1900_Communication_PC".Para.ProduceMode3) AND "DB1042_Timer".HDrillEndTime.Q) OR ((((#HorDrillStep.S20 AND NOT (#HorDrillStep.S22)) OR ((#HorDrillStep.S22 AND NOT (#HorDrillStep.S25)) AND NOT ("DB2500 Visual Chiseling".VisualChiselingMode))) AND "DB1900_Communication_PC".Para.ProduceMode3) AND "DB1042_Timer".GougeTimeOut.Q) OR ((((#HorDrillStep.S20 AND NOT (#HorDrillStep.S22)) OR ((#HorDrillStep.S22 AND NOT (#HorDrillStep.S25)) AND NOT ("DB2500 Visual Chiseling".VisualChiselingMode))) AND "DB1900_Communication_PC".Para.ProduceMode3) AND "DB1042_Timer".CurrentLowTimeOut.Q) OR ((((#HorDrillStep.S20 AND NOT (#HorDrillStep.S22)) OR ((#HorDrillStep.S22 AND NOT (#HorDrillStep.S25)) AND NOT ("DB2500 Visual Chiseling".VisualChiselingMode))) AND "DB1900_Communication_PC".Para.ProduceMode3) AND "DB1042_Timer".CurrentHighTimeOut.Q) OR (((((#HorDrillStep.S20 AND NOT (#HorDrillStep.S22)) OR ((#HorDrillStep.S22 AND NOT (#HorDrillStep.S25)) AND NOT ("DB2500 Visual Chiseling".VisualChiselingMode))) AND "DB1900_Communication_PC".Para.ProduceMode3) AND ("DB1900_Communication_PC".Send.ScrLen >= "DB1900_Communication_PC".Para.DrillDepth))) OR ((((#HorDrillStep.S20 AND NOT (#HorDrillStep.S22)) OR ((#HorDrillStep.S22 AND NOT (#HorDrillStep.S25)) AND NOT ("DB2500 Visual Chiseling".VisualChiselingMode))) AND "DB1900_Communication_PC".Para.ProduceMode3) AND "DB2500 Visual Chiseling".VChiselEndPos) 赋给 #HorDrillStep.GougeStopDrill_End
   #HorDrillStep.GougeStopDrill_End := ((((#HorDrillStep.S20 AND NOT (#HorDrillStep.S22)) OR ((#HorDrillStep.S22 AND NOT (#HorDrillStep.S25)) AND NOT ("DB2500 Visual Chiseling".VisualChiselingMode))) AND "DB1900_Communication_PC".Para.ProduceMode3) AND "DB1042_Timer".HDrillEndTime.Q) OR ((((#HorDrillStep.S20 AND NOT (#HorDrillStep.S22)) OR ((#HorDrillStep.S22 AND NOT (#HorDrillStep.S25)) AND NOT ("DB2500 Visual Chiseling".VisualChiselingMode))) AND "DB1900_Communication_PC".Para.ProduceMode3) AND "DB1042_Timer".GougeTimeOut.Q) OR ((((#HorDrillStep.S20 AND NOT (#HorDrillStep.S22)) OR ((#HorDrillStep.S22 AND NOT (#HorDrillStep.S25)) AND NOT ("DB2500 Visual Chiseling".VisualChiselingMode))) AND "DB1900_Communication_PC".Para.ProduceMode3) AND "DB1042_Timer".CurrentLowTimeOut.Q) OR ((((#HorDrillStep.S20 AND NOT (#HorDrillStep.S22)) OR ((#HorDrillStep.S22 AND NOT (#HorDrillStep.S25)) AND NOT ("DB2500 Visual Chiseling".VisualChiselingMode))) AND "DB1900_Communication_PC".Para.ProduceMode3) AND "DB1042_Timer".CurrentHighTimeOut.Q) OR (((((#HorDrillStep.S20 AND NOT (#HorDrillStep.S22)) OR ((#HorDrillStep.S22 AND NOT (#HorDrillStep.S25)) AND NOT ("DB2500 Visual Chiseling".VisualChiselingMode))) AND "DB1900_Communication_PC".Para.ProduceMode3) AND ("DB1900_Communication_PC".Send.ScrLen >= "DB1900_Communication_PC".Para.DrillDepth))) OR ((((#HorDrillStep.S20 AND NOT (#HorDrillStep.S22)) OR ((#HorDrillStep.S22 AND NOT (#HorDrillStep.S25)) AND NOT ("DB2500 Visual Chiseling".VisualChiselingMode))) AND "DB1900_Communication_PC".Para.ProduceMode3) AND "DB2500 Visual Chiseling".VChiselEndPos);
   // 含义：将 (((((#HorDrillStep.S20 AND NOT (#HorDrillStep.S22)) OR ((#HorDrillStep.S22 AND NOT (#HorDrillStep.S25)) AND NOT ("DB2500 Visual Chiseling".VisualChiselingMode))) AND "DB1900_Communication_PC".Para.ProduceMode3) AND "DB2500 Visual Chiseling".VisualChiselingMode) AND "DB1042_Timer".HDrillEndTime.Q) AND "DB1900_Communication_PC".Para.DrillEndMode 赋给 "DB720_KuKa_MainCtrl".CmdOut.di_VchiselTime_End
   "DB720_KuKa_MainCtrl".CmdOut.di_VchiselTime_End := (((((#HorDrillStep.S20 AND NOT (#HorDrillStep.S22)) OR ((#HorDrillStep.S22 AND NOT (#HorDrillStep.S25)) AND NOT ("DB2500 Visual Chiseling".VisualChiselingMode))) AND "DB1900_Communication_PC".Para.ProduceMode3) AND "DB2500 Visual Chiseling".VisualChiselingMode) AND "DB1042_Timer".HDrillEndTime.Q) AND "DB1900_Communication_PC".Para.DrillEndMode;
   // 含义：将 ((((#HorDrillStep.S20 AND NOT (#HorDrillStep.S22)) OR ((#HorDrillStep.S22 AND NOT (#HorDrillStep.S25)) AND NOT ("DB2500 Visual Chiseling".VisualChiselingMode))) AND #Aux.HDrillOutTime.Q) OR (((((#HorDrillStep.S20 AND NOT (#HorDrillStep.S22)) OR ((#HorDrillStep.S22 AND NOT (#HorDrillStep.S25)) AND NOT ("DB2500 Visual Chiseling".VisualChiselingMode))) AND "DB1042_Timer".CurrentLowTimeOut.Q) OR (((#HorDrillStep.S20 AND NOT (#HorDrillStep.S22)) OR ((#HorDrillStep.S22 AND NOT (#HorDrillStep.S25)) AND NOT ("DB2500 Visual Chiseling".VisualChiselingMode))) AND "DB1042_Timer".CurrentHighTimeOut.Q)) AND NOT (#HorDrillStep.S22)) OR (((((((((#HorDrillStep.S20 AND NOT (#HorDrillStep.S22)) OR ((#HorDrillStep.S22 AND NOT (#HorDrillStep.S25)) AND NOT ("DB2500 Visual Chiseling".VisualChiselingMode))) AND NOT ("DB1900_Communication_PC".Para.ProduceMode3)) AND ("DB1900_Communication_PC".Send.PosNo <= 2))) AND ("DB1900_Communication_PC".Para.DrillWidth <= 28.0))) AND ("DB1900_Communication_PC".Send.ScrLen >= 55.0))) OR (((((#HorDrillStep.S20 AND NOT (#HorDrillStep.S22)) OR ((#HorDrillStep.S22 AND NOT (#HorDrillStep.S25)) AND NOT ("DB2500 Visual Chiseling".VisualChiselingMode))) AND NOT ("DB1900_Communication_PC".Para.ProduceMode3)) AND ("DB1900_Communication_PC".Send.ScrLen >= "DB1900_Communication_PC".Para.DrillDepth))) OR ((((#HorDrillStep.S20 AND NOT (#HorDrillStep.S22)) OR ((#HorDrillStep.S22 AND NOT (#HorDrillStep.S25)) AND NOT ("DB2500 Visual Chiseling".VisualChiselingMode))) AND "DB1042_Timer".HDrillEndTime.Q) AND "DB1900_Communication_PC".Para.DrillEndMode)) AND NOT ("DB1900_Communication_PC".Para.ProduceMode3) 赋给 #HorDrillStep.StopDrill_End
   #HorDrillStep.StopDrill_End := ((((#HorDrillStep.S20 AND NOT (#HorDrillStep.S22)) OR ((#HorDrillStep.S22 AND NOT (#HorDrillStep.S25)) AND NOT ("DB2500 Visual Chiseling".VisualChiselingMode))) AND #Aux.HDrillOutTime.Q) OR (((((#HorDrillStep.S20 AND NOT (#HorDrillStep.S22)) OR ((#HorDrillStep.S22 AND NOT (#HorDrillStep.S25)) AND NOT ("DB2500 Visual Chiseling".VisualChiselingMode))) AND "DB1042_Timer".CurrentLowTimeOut.Q) OR (((#HorDrillStep.S20 AND NOT (#HorDrillStep.S22)) OR ((#HorDrillStep.S22 AND NOT (#HorDrillStep.S25)) AND NOT ("DB2500 Visual Chiseling".VisualChiselingMode))) AND "DB1042_Timer".CurrentHighTimeOut.Q)) AND NOT (#HorDrillStep.S22)) OR (((((((((#HorDrillStep.S20 AND NOT (#HorDrillStep.S22)) OR ((#HorDrillStep.S22 AND NOT (#HorDrillStep.S25)) AND NOT ("DB2500 Visual Chiseling".VisualChiselingMode))) AND NOT ("DB1900_Communication_PC".Para.ProduceMode3)) AND ("DB1900_Communication_PC".Send.PosNo <= 2))) AND ("DB1900_Communication_PC".Para.DrillWidth <= 28.0))) AND ("DB1900_Communication_PC".Send.ScrLen >= 55.0))) OR (((((#HorDrillStep.S20 AND NOT (#HorDrillStep.S22)) OR ((#HorDrillStep.S22 AND NOT (#HorDrillStep.S25)) AND NOT ("DB2500 Visual Chiseling".VisualChiselingMode))) AND NOT ("DB1900_Communication_PC".Para.ProduceMode3)) AND ("DB1900_Communication_PC".Send.ScrLen >= "DB1900_Communication_PC".Para.DrillDepth))) OR ((((#HorDrillStep.S20 AND NOT (#HorDrillStep.S22)) OR ((#HorDrillStep.S22 AND NOT (#HorDrillStep.S25)) AND NOT ("DB2500 Visual Chiseling".VisualChiselingMode))) AND "DB1042_Timer".HDrillEndTime.Q) AND "DB1900_Communication_PC".Para.DrillEndMode)) AND NOT ("DB1900_Communication_PC".Para.ProduceMode3);
   // 含义：条件 (((#HorDrillStep.S20 AND NOT (#HorDrillStep.S22)) OR ((#HorDrillStep.S22 AND NOT (#HorDrillStep.S25)) AND NOT ("DB2500 Visual Chiseling".VisualChiselingMode))) AND TRUE) AND "DB1042_Timer".CurrentLowTimeOut.Q 成立时，将 ("DB1042_Timer".HCLowTimeOutTimes + 1) 传送到 "DB1042_Timer".HCLowTimeOutTimes
   IF (((#HorDrillStep.S20 AND NOT (#HorDrillStep.S22)) OR ((#HorDrillStep.S22 AND NOT (#HorDrillStep.S25)) AND NOT ("DB2500 Visual Chiseling".VisualChiselingMode))) AND TRUE) AND "DB1042_Timer".CurrentLowTimeOut.Q THEN
       "DB1042_Timer".HCLowTimeOutTimes := ("DB1042_Timer".HCLowTimeOutTimes + 1);
   END_IF;
   // 含义：条件 (((#HorDrillStep.S20 AND NOT (#HorDrillStep.S22)) OR ((#HorDrillStep.S22 AND NOT (#HorDrillStep.S25)) AND NOT ("DB2500 Visual Chiseling".VisualChiselingMode))) AND TRUE) AND "DB1042_Timer".CurrentHighTimeOut.Q 成立时，将 ("DB1042_Timer".HCHighTimeOutTimes + 1) 传送到 "DB1042_Timer".HCHighTimeOutTimes
   IF (((#HorDrillStep.S20 AND NOT (#HorDrillStep.S22)) OR ((#HorDrillStep.S22 AND NOT (#HorDrillStep.S25)) AND NOT ("DB2500 Visual Chiseling".VisualChiselingMode))) AND TRUE) AND "DB1042_Timer".CurrentHighTimeOut.Q THEN
       "DB1042_Timer".HCHighTimeOutTimes := ("DB1042_Timer".HCHighTimeOutTimes + 1);
   END_IF;
   // 含义：条件 ((((((((#HorDrillStep.S20 AND NOT (#HorDrillStep.S22)) OR ((#HorDrillStep.S22 AND NOT (#HorDrillStep.S25)) AND NOT ("DB2500 Visual Chiseling".VisualChiselingMode))) AND TRUE) AND #Aux.HDrillOutTime.Q) AND ("DB1900_Communication_PC".Send.ScrLen < "DB1900_Communication_PC".Para.DrillDepth))) AND "DB1900_Communication_PC".Para.ProduceMode3) AND "DB1900_Communication_PC".Para.DrillEndMode) OR (((((((#HorDrillStep.S20 AND NOT (#HorDrillStep.S22)) OR ((#HorDrillStep.S22 AND NOT (#HorDrillStep.S25)) AND NOT ("DB2500 Visual Chiseling".VisualChiselingMode))) AND TRUE) AND #Aux.HDrillOutTime.Q) AND ("DB1900_Communication_PC".Send.ScrLen < "DB1900_Communication_PC".Para.DrillDepth))) AND NOT ("DB1900_Communication_PC".Para.ProduceMode3)) 成立时，将 ("DB1042_Timer".HTimeOutTimes + 1) 传送到 "DB1042_Timer".HTimeOutTimes
   IF ((((((((#HorDrillStep.S20 AND NOT (#HorDrillStep.S22)) OR ((#HorDrillStep.S22 AND NOT (#HorDrillStep.S25)) AND NOT ("DB2500 Visual Chiseling".VisualChiselingMode))) AND TRUE) AND #Aux.HDrillOutTime.Q) AND ("DB1900_Communication_PC".Send.ScrLen < "DB1900_Communication_PC".Para.DrillDepth))) AND "DB1900_Communication_PC".Para.ProduceMode3) AND "DB1900_Communication_PC".Para.DrillEndMode) OR (((((((#HorDrillStep.S20 AND NOT (#HorDrillStep.S22)) OR ((#HorDrillStep.S22 AND NOT (#HorDrillStep.S25)) AND NOT ("DB2500 Visual Chiseling".VisualChiselingMode))) AND TRUE) AND #Aux.HDrillOutTime.Q) AND ("DB1900_Communication_PC".Send.ScrLen < "DB1900_Communication_PC".Para.DrillDepth))) AND NOT ("DB1900_Communication_PC".Para.ProduceMode3)) THEN
       "DB1042_Timer".HTimeOutTimes := ("DB1042_Timer".HTimeOutTimes + 1);
   END_IF;
   // 含义：条件 (((((#HorDrillStep.S20 AND NOT (#HorDrillStep.S22)) OR ((#HorDrillStep.S22 AND NOT (#HorDrillStep.S25)) AND NOT ("DB2500 Visual Chiseling".VisualChiselingMode))) AND TRUE) AND ("DB1042_Timer".HCLowTimeOutTimes > 2))) AND NOT ("DB1900_Communication_PC".Para.ProduceMode3) 成立时，将 TRUE 传送到 "DB1148_PromptBeeper".Public.CurrentLowTimeOut
   IF (((((#HorDrillStep.S20 AND NOT (#HorDrillStep.S22)) OR ((#HorDrillStep.S22 AND NOT (#HorDrillStep.S25)) AND NOT ("DB2500 Visual Chiseling".VisualChiselingMode))) AND TRUE) AND ("DB1042_Timer".HCLowTimeOutTimes > 2))) AND NOT ("DB1900_Communication_PC".Para.ProduceMode3) THEN
       "DB1148_PromptBeeper".Public.CurrentLowTimeOut := TRUE;
   END_IF;
   // 含义：条件 (((((#HorDrillStep.S20 AND NOT (#HorDrillStep.S22)) OR ((#HorDrillStep.S22 AND NOT (#HorDrillStep.S25)) AND NOT ("DB2500 Visual Chiseling".VisualChiselingMode))) AND TRUE) AND ("DB1042_Timer".HCLowTimeOutTimes > 2))) AND NOT ("DB1900_Communication_PC".Para.ProduceMode3) 成立时，将 TRUE 传送到 #HorDrillStep.ErrEnd
   IF (((((#HorDrillStep.S20 AND NOT (#HorDrillStep.S22)) OR ((#HorDrillStep.S22 AND NOT (#HorDrillStep.S25)) AND NOT ("DB2500 Visual Chiseling".VisualChiselingMode))) AND TRUE) AND ("DB1042_Timer".HCLowTimeOutTimes > 2))) AND NOT ("DB1900_Communication_PC".Para.ProduceMode3) THEN
       #HorDrillStep.ErrEnd := TRUE;
   END_IF;
   // 含义：条件 (((((#HorDrillStep.S20 AND NOT (#HorDrillStep.S22)) OR ((#HorDrillStep.S22 AND NOT (#HorDrillStep.S25)) AND NOT ("DB2500 Visual Chiseling".VisualChiselingMode))) AND TRUE) AND ("DB1042_Timer".HCLowTimeOutTimes > 2))) AND NOT ("DB1900_Communication_PC".Para.ProduceMode3) 成立时，将 0 传送到 "DB1042_Timer".HCLowTimeOutTimes
   IF (((((#HorDrillStep.S20 AND NOT (#HorDrillStep.S22)) OR ((#HorDrillStep.S22 AND NOT (#HorDrillStep.S25)) AND NOT ("DB2500 Visual Chiseling".VisualChiselingMode))) AND TRUE) AND ("DB1042_Timer".HCLowTimeOutTimes > 2))) AND NOT ("DB1900_Communication_PC".Para.ProduceMode3) THEN
       "DB1042_Timer".HCLowTimeOutTimes := 0;
   END_IF;
   // 含义：条件 ((((((#HorDrillStep.S20 AND NOT (#HorDrillStep.S22)) OR ((#HorDrillStep.S22 AND NOT (#HorDrillStep.S25)) AND NOT ("DB2500 Visual Chiseling".VisualChiselingMode))) AND TRUE) AND NOT ("DB1900_Communication_PC".Para.ProduceMode3)) AND ("DB1042_Timer".HCHighTimeOutTimes > 2))) OR ((((((#HorDrillStep.S20 AND NOT (#HorDrillStep.S22)) OR ((#HorDrillStep.S22 AND NOT (#HorDrillStep.S25)) AND NOT ("DB2500 Visual Chiseling".VisualChiselingMode))) AND TRUE) AND "DB1900_Communication_PC".Para.ProduceMode3) AND ("DB1042_Timer".HCLowTimeOutTimes >= 5))) 成立时，将 TRUE 传送到 "DB1148_PromptBeeper".Public.CurrentHighTimeOut
   IF ((((((#HorDrillStep.S20 AND NOT (#HorDrillStep.S22)) OR ((#HorDrillStep.S22 AND NOT (#HorDrillStep.S25)) AND NOT ("DB2500 Visual Chiseling".VisualChiselingMode))) AND TRUE) AND NOT ("DB1900_Communication_PC".Para.ProduceMode3)) AND ("DB1042_Timer".HCHighTimeOutTimes > 2))) OR ((((((#HorDrillStep.S20 AND NOT (#HorDrillStep.S22)) OR ((#HorDrillStep.S22 AND NOT (#HorDrillStep.S25)) AND NOT ("DB2500 Visual Chiseling".VisualChiselingMode))) AND TRUE) AND "DB1900_Communication_PC".Para.ProduceMode3) AND ("DB1042_Timer".HCLowTimeOutTimes >= 5))) THEN
       "DB1148_PromptBeeper".Public.CurrentHighTimeOut := TRUE;
   END_IF;
   // 含义：条件 ((((((#HorDrillStep.S20 AND NOT (#HorDrillStep.S22)) OR ((#HorDrillStep.S22 AND NOT (#HorDrillStep.S25)) AND NOT ("DB2500 Visual Chiseling".VisualChiselingMode))) AND TRUE) AND NOT ("DB1900_Communication_PC".Para.ProduceMode3)) AND ("DB1042_Timer".HCHighTimeOutTimes > 2))) OR ((((((#HorDrillStep.S20 AND NOT (#HorDrillStep.S22)) OR ((#HorDrillStep.S22 AND NOT (#HorDrillStep.S25)) AND NOT ("DB2500 Visual Chiseling".VisualChiselingMode))) AND TRUE) AND "DB1900_Communication_PC".Para.ProduceMode3) AND ("DB1042_Timer".HCLowTimeOutTimes >= 5))) 成立时，将 TRUE 传送到 #HorDrillStep.ErrEnd
   IF ((((((#HorDrillStep.S20 AND NOT (#HorDrillStep.S22)) OR ((#HorDrillStep.S22 AND NOT (#HorDrillStep.S25)) AND NOT ("DB2500 Visual Chiseling".VisualChiselingMode))) AND TRUE) AND NOT ("DB1900_Communication_PC".Para.ProduceMode3)) AND ("DB1042_Timer".HCHighTimeOutTimes > 2))) OR ((((((#HorDrillStep.S20 AND NOT (#HorDrillStep.S22)) OR ((#HorDrillStep.S22 AND NOT (#HorDrillStep.S25)) AND NOT ("DB2500 Visual Chiseling".VisualChiselingMode))) AND TRUE) AND "DB1900_Communication_PC".Para.ProduceMode3) AND ("DB1042_Timer".HCLowTimeOutTimes >= 5))) THEN
       #HorDrillStep.ErrEnd := TRUE;
   END_IF;
   // 含义：条件 ((((((#HorDrillStep.S20 AND NOT (#HorDrillStep.S22)) OR ((#HorDrillStep.S22 AND NOT (#HorDrillStep.S25)) AND NOT ("DB2500 Visual Chiseling".VisualChiselingMode))) AND TRUE) AND NOT ("DB1900_Communication_PC".Para.ProduceMode3)) AND ("DB1042_Timer".HCHighTimeOutTimes > 2))) OR ((((((#HorDrillStep.S20 AND NOT (#HorDrillStep.S22)) OR ((#HorDrillStep.S22 AND NOT (#HorDrillStep.S25)) AND NOT ("DB2500 Visual Chiseling".VisualChiselingMode))) AND TRUE) AND "DB1900_Communication_PC".Para.ProduceMode3) AND ("DB1042_Timer".HCLowTimeOutTimes >= 5))) 成立时，将 0 传送到 "DB1042_Timer".HCHighTimeOutTimes
   IF ((((((#HorDrillStep.S20 AND NOT (#HorDrillStep.S22)) OR ((#HorDrillStep.S22 AND NOT (#HorDrillStep.S25)) AND NOT ("DB2500 Visual Chiseling".VisualChiselingMode))) AND TRUE) AND NOT ("DB1900_Communication_PC".Para.ProduceMode3)) AND ("DB1042_Timer".HCHighTimeOutTimes > 2))) OR ((((((#HorDrillStep.S20 AND NOT (#HorDrillStep.S22)) OR ((#HorDrillStep.S22 AND NOT (#HorDrillStep.S25)) AND NOT ("DB2500 Visual Chiseling".VisualChiselingMode))) AND TRUE) AND "DB1900_Communication_PC".Para.ProduceMode3) AND ("DB1042_Timer".HCLowTimeOutTimes >= 5))) THEN
       "DB1042_Timer".HCHighTimeOutTimes := 0;
   END_IF;
   // 含义：条件 (((((#HorDrillStep.S20 AND NOT (#HorDrillStep.S22)) OR ((#HorDrillStep.S22 AND NOT (#HorDrillStep.S25)) AND NOT ("DB2500 Visual Chiseling".VisualChiselingMode))) AND TRUE) AND NOT ("DB1900_Communication_PC".Para.ProduceMode3)) AND ("DB1900_Communication_PC".Send.ScrLen >= #Aux.DrillDepthMax)) 成立时，将 TRUE 传送到 "DB1148_PromptBeeper".Public.DrillDepthErr
   IF (((((#HorDrillStep.S20 AND NOT (#HorDrillStep.S22)) OR ((#HorDrillStep.S22 AND NOT (#HorDrillStep.S25)) AND NOT ("DB2500 Visual Chiseling".VisualChiselingMode))) AND TRUE) AND NOT ("DB1900_Communication_PC".Para.ProduceMode3)) AND ("DB1900_Communication_PC".Send.ScrLen >= #Aux.DrillDepthMax)) THEN
       "DB1148_PromptBeeper".Public.DrillDepthErr := TRUE;
   END_IF;
   // 含义：条件 (((((((((#HorDrillStep.S20 AND NOT (#HorDrillStep.S22)) OR ((#HorDrillStep.S22 AND NOT (#HorDrillStep.S25)) AND NOT ("DB2500 Visual Chiseling".VisualChiselingMode))) AND "DB720_KuKa_MainCtrl".StatusIn.do_HorDril_Pos) OR (((#HorDrillStep.S20 AND NOT (#HorDrillStep.S22)) OR ((#HorDrillStep.S22 AND NOT (#HorDrillStep.S25)) AND NOT ("DB2500 Visual Chiseling".VisualChiselingMode))) AND "DB720_KuKa_MainCtrl".StatusIn.do_Gouge_Pos)) AND NOT (#HorDrillStep.StopDrill_Ack)) AND ("DB1900_Communication_PC".Recv.Current_2 > "DB1900_Communication_PC".Para.CurrentMinLimit))) AND ("DB1900_Communication_PC".Recv.Current_2 < "DB1900_Communication_PC".Para.CurrentMaxLimit))) AND "DB1042_Timer".HCurrentLastTime.Q 成立时，将 0 传送到 "DB1042_Timer".HCLowTimeOutTimes
   IF (((((((((#HorDrillStep.S20 AND NOT (#HorDrillStep.S22)) OR ((#HorDrillStep.S22 AND NOT (#HorDrillStep.S25)) AND NOT ("DB2500 Visual Chiseling".VisualChiselingMode))) AND "DB720_KuKa_MainCtrl".StatusIn.do_HorDril_Pos) OR (((#HorDrillStep.S20 AND NOT (#HorDrillStep.S22)) OR ((#HorDrillStep.S22 AND NOT (#HorDrillStep.S25)) AND NOT ("DB2500 Visual Chiseling".VisualChiselingMode))) AND "DB720_KuKa_MainCtrl".StatusIn.do_Gouge_Pos)) AND NOT (#HorDrillStep.StopDrill_Ack)) AND ("DB1900_Communication_PC".Recv.Current_2 > "DB1900_Communication_PC".Para.CurrentMinLimit))) AND ("DB1900_Communication_PC".Recv.Current_2 < "DB1900_Communication_PC".Para.CurrentMaxLimit))) AND "DB1042_Timer".HCurrentLastTime.Q THEN
       "DB1042_Timer".HCLowTimeOutTimes := 0;
   END_IF;
   // 含义：调用计数器实例 "DB1042_Timer".HCurrentLastTime.TON（上升沿计数，当前值写入 CV）
   "DB1042_Timer".HCurrentLastTime.TON(IN := ((((((((#HorDrillStep.S20 AND NOT (#HorDrillStep.S22)) OR ((#HorDrillStep.S22 AND NOT (#HorDrillStep.S25)) AND NOT ("DB2500 Visual Chiseling".VisualChiselingMode))) AND "DB720_KuKa_MainCtrl".StatusIn.do_HorDril_Pos) OR (((#HorDrillStep.S20 AND NOT (#HorDrillStep.S22)) OR ((#HorDrillStep.S22 AND NOT (#HorDrillStep.S25)) AND NOT ("DB2500 Visual Chiseling".VisualChiselingMode))) AND "DB720_KuKa_MainCtrl".StatusIn.do_Gouge_Pos)) AND NOT (#HorDrillStep.StopDrill_Ack)) AND ("DB1900_Communication_PC".Recv.Current_2 > "DB1900_Communication_PC".Para.CurrentMinLimit))) AND ("DB1900_Communication_PC".Recv.Current_2 < "DB1900_Communication_PC".Para.CurrentMaxLimit)),
                                       PT := T#500ms);
   // 含义：条件 ((((((((#HorDrillStep.S20 AND NOT (#HorDrillStep.S22)) OR ((#HorDrillStep.S22 AND NOT (#HorDrillStep.S25)) AND NOT ("DB2500 Visual Chiseling".VisualChiselingMode))) AND "DB720_KuKa_MainCtrl".StatusIn.do_HorDril_Pos) OR (((#HorDrillStep.S20 AND NOT (#HorDrillStep.S22)) OR ((#HorDrillStep.S22 AND NOT (#HorDrillStep.S25)) AND NOT ("DB2500 Visual Chiseling".VisualChiselingMode))) AND "DB720_KuKa_MainCtrl".StatusIn.do_Gouge_Pos)) AND #HorDrillStep.StopDrill_Ack) AND NOT ("DB1900_Communication_PC".Para.ProduceMode3)) AND ("DB1900_Communication_PC".Send.ScrLen >= #Aux.DrillDepthMin))) OR (((((((#HorDrillStep.S20 AND NOT (#HorDrillStep.S22)) OR ((#HorDrillStep.S22 AND NOT (#HorDrillStep.S25)) AND NOT ("DB2500 Visual Chiseling".VisualChiselingMode))) AND "DB720_KuKa_MainCtrl".StatusIn.do_HorDril_Pos) OR (((#HorDrillStep.S20 AND NOT (#HorDrillStep.S22)) OR ((#HorDrillStep.S22 AND NOT (#HorDrillStep.S25)) AND NOT ("DB2500 Visual Chiseling".VisualChiselingMode))) AND "DB720_KuKa_MainCtrl".StatusIn.do_Gouge_Pos)) AND #HorDrillStep.StopDrill_Ack) AND "DB1042_Timer".HDrillEndTime.Q) AND "DB1900_Communication_PC".Para.DrillEndMode) 成立时，将 0 传送到 "DB1042_Timer".HTimeOutTimes
   IF ((((((((#HorDrillStep.S20 AND NOT (#HorDrillStep.S22)) OR ((#HorDrillStep.S22 AND NOT (#HorDrillStep.S25)) AND NOT ("DB2500 Visual Chiseling".VisualChiselingMode))) AND "DB720_KuKa_MainCtrl".StatusIn.do_HorDril_Pos) OR (((#HorDrillStep.S20 AND NOT (#HorDrillStep.S22)) OR ((#HorDrillStep.S22 AND NOT (#HorDrillStep.S25)) AND NOT ("DB2500 Visual Chiseling".VisualChiselingMode))) AND "DB720_KuKa_MainCtrl".StatusIn.do_Gouge_Pos)) AND #HorDrillStep.StopDrill_Ack) AND NOT ("DB1900_Communication_PC".Para.ProduceMode3)) AND ("DB1900_Communication_PC".Send.ScrLen >= #Aux.DrillDepthMin))) OR (((((((#HorDrillStep.S20 AND NOT (#HorDrillStep.S22)) OR ((#HorDrillStep.S22 AND NOT (#HorDrillStep.S25)) AND NOT ("DB2500 Visual Chiseling".VisualChiselingMode))) AND "DB720_KuKa_MainCtrl".StatusIn.do_HorDril_Pos) OR (((#HorDrillStep.S20 AND NOT (#HorDrillStep.S22)) OR ((#HorDrillStep.S22 AND NOT (#HorDrillStep.S25)) AND NOT ("DB2500 Visual Chiseling".VisualChiselingMode))) AND "DB720_KuKa_MainCtrl".StatusIn.do_Gouge_Pos)) AND #HorDrillStep.StopDrill_Ack) AND "DB1042_Timer".HDrillEndTime.Q) AND "DB1900_Communication_PC".Para.DrillEndMode) THEN
       "DB1042_Timer".HTimeOutTimes := 0;
   END_IF;
   // 含义：条件 ((#HorDrillStep.S20 AND NOT (#HorDrillStep.S22)) OR ((#HorDrillStep.S22 AND NOT (#HorDrillStep.S25)) AND NOT ("DB2500 Visual Chiseling".VisualChiselingMode))) AND "DB1042_Timer".FixtureStuckTimeOut.Q 成立时，将 TRUE 传送到 #HorDrillStep.ErrEnd
   IF ((#HorDrillStep.S20 AND NOT (#HorDrillStep.S22)) OR ((#HorDrillStep.S22 AND NOT (#HorDrillStep.S25)) AND NOT ("DB2500 Visual Chiseling".VisualChiselingMode))) AND "DB1042_Timer".FixtureStuckTimeOut.Q THEN
       #HorDrillStep.ErrEnd := TRUE;
   END_IF;
   // 含义：条件 ((#HorDrillStep.S20 AND NOT (#HorDrillStep.S22)) OR ((#HorDrillStep.S22 AND NOT (#HorDrillStep.S25)) AND NOT ("DB2500 Visual Chiseling".VisualChiselingMode))) AND "DB1042_Timer".FixtureStuckTimeOut.Q 成立时，将 TRUE 传送到 "DB1148_PromptBeeper".Public.BitStuckErr_Fixture
   IF ((#HorDrillStep.S20 AND NOT (#HorDrillStep.S22)) OR ((#HorDrillStep.S22 AND NOT (#HorDrillStep.S25)) AND NOT ("DB2500 Visual Chiseling".VisualChiselingMode))) AND "DB1042_Timer".FixtureStuckTimeOut.Q THEN
       "DB1148_PromptBeeper".Public.BitStuckErr_Fixture := TRUE;
   END_IF;
   // 含义：条件 ((#HorDrillStep.S20 AND NOT (#HorDrillStep.S22)) OR ((#HorDrillStep.S22 AND NOT (#HorDrillStep.S25)) AND NOT ("DB2500 Visual Chiseling".VisualChiselingMode))) AND "DB1042_Timer".DrillingHighCurrentOut.Q 成立时，将 TRUE 传送到 #HorDrillStep.ErrEnd
   IF ((#HorDrillStep.S20 AND NOT (#HorDrillStep.S22)) OR ((#HorDrillStep.S22 AND NOT (#HorDrillStep.S25)) AND NOT ("DB2500 Visual Chiseling".VisualChiselingMode))) AND "DB1042_Timer".DrillingHighCurrentOut.Q THEN
       #HorDrillStep.ErrEnd := TRUE;
   END_IF;
   // 含义：条件 ((#HorDrillStep.S20 AND NOT (#HorDrillStep.S22)) OR ((#HorDrillStep.S22 AND NOT (#HorDrillStep.S25)) AND NOT ("DB2500 Visual Chiseling".VisualChiselingMode))) AND "DB1042_Timer".DrillingHighCurrentOut.Q 成立时，将 TRUE 传送到 "DB1148_PromptBeeper".Public.BitStuckErr_HighCurrent
   IF ((#HorDrillStep.S20 AND NOT (#HorDrillStep.S22)) OR ((#HorDrillStep.S22 AND NOT (#HorDrillStep.S25)) AND NOT ("DB2500 Visual Chiseling".VisualChiselingMode))) AND "DB1042_Timer".DrillingHighCurrentOut.Q THEN
       "DB1148_PromptBeeper".Public.BitStuckErr_HighCurrent := TRUE;
   END_IF;

   // ---------- 网络 21 ----------
   // 标题：TaskDone
   // 含义：条件 ((#HorDrillStep.S25 OR (#HorDrillStep.S22 AND "DB2500 Visual Chiseling".VisualChiselingMode) OR #HorDrillStep.ErrEnd OR #HorDrillStep.ByPass) AND NOT (#HorDrillStep.S27)) AND NOT (#HorDrillStep.ErrEnd) 成立时，将 TRUE 传送到 #HorDrillStep.TaskIO
   IF ((#HorDrillStep.S25 OR (#HorDrillStep.S22 AND "DB2500 Visual Chiseling".VisualChiselingMode) OR #HorDrillStep.ErrEnd OR #HorDrillStep.ByPass) AND NOT (#HorDrillStep.S27)) AND NOT (#HorDrillStep.ErrEnd) THEN
       #HorDrillStep.TaskIO := TRUE;
   END_IF;
   // 含义：条件 ((#HorDrillStep.S25 OR (#HorDrillStep.S22 AND "DB2500 Visual Chiseling".VisualChiselingMode) OR #HorDrillStep.ErrEnd OR #HorDrillStep.ByPass) AND NOT (#HorDrillStep.S27)) AND #HorDrillStep.ErrEnd 成立时，将 TRUE 传送到 #HorDrillStep.TaskNIO
   IF ((#HorDrillStep.S25 OR (#HorDrillStep.S22 AND "DB2500 Visual Chiseling".VisualChiselingMode) OR #HorDrillStep.ErrEnd OR #HorDrillStep.ByPass) AND NOT (#HorDrillStep.S27)) AND #HorDrillStep.ErrEnd THEN
       #HorDrillStep.TaskNIO := TRUE;
   END_IF;
   // 含义：条件 (#HorDrillStep.S25 OR (#HorDrillStep.S22 AND "DB2500 Visual Chiseling".VisualChiselingMode) OR #HorDrillStep.ErrEnd OR #HorDrillStep.ByPass) AND NOT (#HorDrillStep.S27) 成立时，将 FALSE 传送到 "DB1042_Timer".FirstStart
   IF (#HorDrillStep.S25 OR (#HorDrillStep.S22 AND "DB2500 Visual Chiseling".VisualChiselingMode) OR #HorDrillStep.ErrEnd OR #HorDrillStep.ByPass) AND NOT (#HorDrillStep.S27) THEN
       "DB1042_Timer".FirstStart := FALSE;
   END_IF;
   // 含义：将 #HorDrillStep.S25 OR (#HorDrillStep.S22 AND "DB2500 Visual Chiseling".VisualChiselingMode) OR #HorDrillStep.ErrEnd OR #HorDrillStep.ByPass 赋给 #HorDrillStep.S27
   #HorDrillStep.S27 := #HorDrillStep.S25 OR (#HorDrillStep.S22 AND "DB2500 Visual Chiseling".VisualChiselingMode) OR #HorDrillStep.ErrEnd OR #HorDrillStep.ByPass;

   // ---------- 网络 22 ----------
   // 标题：结束
   // 注释：Added DB2700.VisualChiselingEnd  by WXY, 20220615.
   // 含义：将 #HorDrillStep.S27 AND NOT (#HorDrillStep.StartCmd) 赋给 #HorDrillStep.StepEnd
   #HorDrillStep.StepEnd := #HorDrillStep.S27 AND NOT (#HorDrillStep.StartCmd);
   // 含义：条件 #HorDrillStep.S27 AND #HorDrillStep.ErrEnd 成立时，将 TRUE 传送到 "DB1080_Component".Robot.Cmd.Auto.Stop
   IF #HorDrillStep.S27 AND #HorDrillStep.ErrEnd THEN
       "DB1080_Component".Robot.Cmd.Auto.Stop := TRUE;
   END_IF;
   // 含义：将 (#HorDrillStep.S27 AND "DB1080_Component".Robot.Status.TaskDone) OR (#HorDrillStep.S27 AND #HorDrillStep.TaskDone) 赋给 #HorDrillStep.TaskDone
   #HorDrillStep.TaskDone := (#HorDrillStep.S27 AND "DB1080_Component".Robot.Status.TaskDone) OR (#HorDrillStep.S27 AND #HorDrillStep.TaskDone);
   // 含义：条件 (((#HorDrillStep.S27 AND "DB1080_Component".Robot.Status.TaskDone) OR (#HorDrillStep.S27 AND #HorDrillStep.TaskDone)) AND "DB1900_Communication_PC".Para.ProduceMode3) AND "DB2500 Visual Chiseling".VisualChiselingMode 成立时，将 FALSE 传送到 "DB2500 Visual Chiseling".VisualChiselingStart
   IF (((#HorDrillStep.S27 AND "DB1080_Component".Robot.Status.TaskDone) OR (#HorDrillStep.S27 AND #HorDrillStep.TaskDone)) AND "DB1900_Communication_PC".Para.ProduceMode3) AND "DB2500 Visual Chiseling".VisualChiselingMode THEN
       "DB2500 Visual Chiseling".VisualChiselingStart := FALSE;
   END_IF;
   // 含义：条件 (((#HorDrillStep.S27 AND "DB1080_Component".Robot.Status.TaskDone) OR (#HorDrillStep.S27 AND #HorDrillStep.TaskDone)) AND "DB1900_Communication_PC".Para.ProduceMode3) AND "DB2500 Visual Chiseling".VisualChiselingMode 成立时，将 TRUE 传送到 "DB2500 Visual Chiseling".VisualChiselingEnd
   IF (((#HorDrillStep.S27 AND "DB1080_Component".Robot.Status.TaskDone) OR (#HorDrillStep.S27 AND #HorDrillStep.TaskDone)) AND "DB1900_Communication_PC".Para.ProduceMode3) AND "DB2500 Visual Chiseling".VisualChiselingMode THEN
       "DB2500 Visual Chiseling".VisualChiselingEnd := TRUE;
   END_IF;

   // ---------- 网络 23 ----------
   // 含义：将 FALSE 赋给 #HorDrillStep.StartCmd
   #HorDrillStep.StartCmd := FALSE;
   // 含义：条件 ("DB1900_Communication_PC".Para.ProduceMode3 AND NOT ("DB720_KuKa_MainCtrl".StatusIn.do_DrilEnd_Pos)) AND NOT ("DB2600 FT Control".FTControlBreak) 成立时，将 FALSE 传送到 "DB2500 Visual Chiseling".VChiselEndPos
   IF ("DB1900_Communication_PC".Para.ProduceMode3 AND NOT ("DB720_KuKa_MainCtrl".StatusIn.do_DrilEnd_Pos)) AND NOT ("DB2600 FT Control".FTControlBreak) THEN
       "DB2500 Visual Chiseling".VChiselEndPos := FALSE;
   END_IF;
   // 含义：条件 "ManMode_M" AND "ErrRst_M" 成立时，将 FALSE 传送到 "DB1148_PromptBeeper".Public.HorChiselStuckErr
   IF "ManMode_M" AND "ErrRst_M" THEN
       "DB1148_PromptBeeper".Public.HorChiselStuckErr := FALSE;
   END_IF;

   // ---------- 网络 24 ----------
   // （空白网络）
END_FUNCTION_BLOCK

FUNCTION_BLOCK "FB1063_DownDrillAutoStep"   // FB1063, SCL
{ S7_Optimized_Access := 'TRUE' }
// ============================================================
//  Block: FB1063_DownDrillAutoStep
//  ============================================================
//  编号：FB1063
//  原始语言：LAD（规则翻译为 SCL）
//  含义：PosNo is ToolNo, not HoleNo.
   VAR
      Aux : Struct   // 静态变量
         StartDrill : Bool;   // 静态变量
         DrillDepthMid : DInt;   // 打孔深度中间变量
         DrillDepthMax : Real;   // 静态变量
         DrillDepthMin : Real;   // 静态变量
         DDrillTime : IEC_TIMER;   // 静态变量
      END_STRUCT;
      EdgeDetc : Struct   // 静态变量
         Pulse : Array[0..15] of Bool;   // 静态变量
      END_STRUCT;
      DownDrillStep : Struct   // 向下钻孔
         Busy : Bool;   // 静态变量
         StartCmd : Bool;   // 静态变量
         OKToStart : Bool;   // 静态变量
         TaskDone : Bool;   // 静态变量
         StepStart : Bool;   // 静态变量
         StepEnd : Bool;   // 静态变量
         ErrEnd : Bool;   // 静态变量
         ByPass : Bool;   // 静态变量
         TaskIO : Bool;   // 静态变量
         TaskNIO : Bool;   // 静态变量
         S1 : Bool;   // 静态变量
         S2 : Bool;   // 静态变量
         S3 : Bool;   // 静态变量
         S4 : Bool;   // 静态变量
         S5 : Bool;   // 静态变量
         S6 : Bool;   // 静态变量
         S7 : Bool;   // 静态变量
         S8 : Bool;   // 静态变量
         S9 : Bool;   // 静态变量
         S10 : Bool;   // 静态变量
         S11 : Bool;   // 静态变量
         S12 : Bool;   // 静态变量
         S13 : Bool;   // 静态变量
         S14 : Bool;   // 静态变量
         S15 : Bool;   // 静态变量
         S16 : Bool;   // 静态变量
         S17 : Bool;   // 静态变量
         S18 : Bool;   // 静态变量
         S19 : Bool;   // 静态变量
         S20 : Bool;   // 静态变量
         S21 : Bool;   // 静态变量
         S22 : Bool;   // 静态变量
         S23 : Bool;   // 静态变量
         S24 : Bool;   // 静态变量
         S25 : Bool;   // 静态变量
         S26 : Bool;   // 静态变量
         S27 : Bool;   // 静态变量
         S28 : Bool;   // 静态变量
         S29 : Bool;   // 静态变量
         S30 : Bool;   // 静态变量
         S31 : Bool;   // 静态变量
         S32 : Bool;   // 静态变量
         S33 : Bool;   // 静态变量
         S34 : Bool;   // 静态变量
         S35 : Bool;   // 静态变量
         S36 : Bool;   // 静态变量
         S37 : Bool;   // 静态变量
         S38 : Bool;   // 静态变量
         S39 : Bool;   // 静态变量
         S40 : Bool;   // 静态变量
         S41 : Bool;   // 静态变量
         S42 : Bool;   // 静态变量
         S43 : Bool;   // 静态变量
         S44 : Bool;   // 静态变量
         S45 : Bool;   // 静态变量
         S46 : Bool;   // 静态变量
         S47 : Bool;   // 静态变量
         S48 : Bool;   // 静态变量
         S49 : Bool;   // 静态变量
         S50 : Bool;   // 静态变量
         S51 : Bool;   // 静态变量
         S52 : Bool;   // 静态变量
         S53 : Bool;   // 静态变量
         S54 : Bool;   // 静态变量
         S55 : Bool;   // 静态变量
         S56 : Bool;   // 静态变量
         S57 : Bool;   // 静态变量
         S58 : Bool;   // 静态变量
         S59 : Bool;   // 静态变量
         S60 : Bool;   // 静态变量
         S61 : Bool;   // 静态变量
         S62 : Bool;   // 静态变量
         S63 : Bool;   // 静态变量
         S64 : Bool;   // 静态变量
         S65 : Bool;   // 静态变量
         InitForcePulse : Bool;   // 静态变量
         ChiselEndPos : Bool;   // 静态变量
         StopDrill_Ack : Bool;   // 静态变量
         StopDrill_End : Bool;   // 静态变量
      END_STRUCT;
      PT : Time;   // 静态变量
      ET : Time;   // 静态变量
      IN : Bool;   // 静态变量
      Q : Bool;   // 静态变量
   END_VAR
   VAR_TEMP
      DownPosMod : Int;   // 临时变量
   END_VAR
BEGIN

   // ---------- 网络 1 ----------
   // （空白网络）

   // ---------- 网络 2 ----------
   // 标题：********************************垂直向下钻孔Start**************************************
   // 含义：将 (("DB720_KuKa_MainCtrl".Ctrl_Out.RobotAction = 0) AND "DB720_KuKa_MainCtrl".Aux.ToolAtPos) AND NOT ("DB1148_PromptBeeper".Public.RobotNotReady) 赋给 #DownDrillStep.OKToStart
   #DownDrillStep.OKToStart := (("DB720_KuKa_MainCtrl".Ctrl_Out.RobotAction = 0) AND "DB720_KuKa_MainCtrl".Aux.ToolAtPos) AND NOT ("DB1148_PromptBeeper".Public.RobotNotReady);
   // 含义：条件 (("ManMode_M" AND "DB1900_Communication_PC".Recv.RobotDrillTPPB) AND ("DB1900_Communication_PC".Recv.ChooseProgNo = 2)) 成立时，将 TRUE 传送到 #DownDrillStep.StartCmd
   IF (("ManMode_M" AND "DB1900_Communication_PC".Recv.RobotDrillTPPB) AND ("DB1900_Communication_PC".Recv.ChooseProgNo = 2)) THEN
       #DownDrillStep.StartCmd := TRUE;
   END_IF;
   // 含义：条件 "DB1060_AutoStep".DownDrillAutoStep.DownDrillStep.StepStart AND "DB1900_Communication_PC".Para.ProduceMode3 成立时，将 ("DB1900_Communication_PC".Para.DrillDepth + 0.0) 传送到 #Aux.DrillDepthMid
   IF "DB1060_AutoStep".DownDrillAutoStep.DownDrillStep.StepStart AND "DB1900_Communication_PC".Para.ProduceMode3 THEN
       #Aux.DrillDepthMid := ("DB1900_Communication_PC".Para.DrillDepth + 0.0);
   END_IF;
   // 含义：将 SWAP(#Aux.DrillDepthMid) 赋给 "DB720_KuKa_MainCtrl".CmdOut.gi_Depth
   "DB720_KuKa_MainCtrl".CmdOut.gi_Depth := SWAP(#Aux.DrillDepthMid);
   // 含义：条件 "DB1060_AutoStep".DownDrillAutoStep.DownDrillStep.StepStart AND "DB1900_Communication_PC".Para.ProduceMode3 成立时，将 "DB1910_DrillData".AUX.LayerNo 传送到 "DB720_KuKa_MainCtrl".CmdOut.gi_LayerNum
   IF "DB1060_AutoStep".DownDrillAutoStep.DownDrillStep.StepStart AND "DB1900_Communication_PC".Para.ProduceMode3 THEN
       "DB720_KuKa_MainCtrl".CmdOut.gi_LayerNum := "DB1910_DrillData".AUX.LayerNo;
   END_IF;
   // 含义：条件 "DB1060_AutoStep".DownDrillAutoStep.DownDrillStep.StepStart AND NOT ("DB1900_Communication_PC".Para.ProduceMode3) 成立时，将 ("DB1900_Communication_PC".Para.DrillDepth + 5.0) 传送到 #Aux.DrillDepthMid
   IF "DB1060_AutoStep".DownDrillAutoStep.DownDrillStep.StepStart AND NOT ("DB1900_Communication_PC".Para.ProduceMode3) THEN
       #Aux.DrillDepthMid := ("DB1900_Communication_PC".Para.DrillDepth + 5.0);
   END_IF;
   // 含义：将 SWAP(#Aux.DrillDepthMid) 赋给 "DB720_KuKa_MainCtrl".CmdOut.gi_Depth
   "DB720_KuKa_MainCtrl".CmdOut.gi_Depth := SWAP(#Aux.DrillDepthMid);

   // ---------- 网络 3 ----------
   // 标题：*******************************打孔超时计时****************************************
   // 含义：调用定时器实例 #Aux.DDrillTime.TON
   #Aux.DDrillTime.TON(IN := "DB720_KuKa_MainCtrl".StatusIn.do_DownDril_Pos AND NOT ("DB1148_PromptBeeper".Public.DrillTimeOut),
                       PT := "DB1900_Communication_PC".Para.TimeOut);

   // ---------- 网络 4 ----------
   // 标题：**********************************钻孔区间*******************************************
   // 含义：将 ("DB1900_Communication_PC".Para.DrillDepth + 10.0) 赋给 #Aux.DrillDepthMax
   #Aux.DrillDepthMax := ("DB1900_Communication_PC".Para.DrillDepth + 10.0);
   // 含义：将 ("DB1900_Communication_PC".Para.DrillDepth - 5.0) 赋给 #Aux.DrillDepthMin
   #Aux.DrillDepthMin := ("DB1900_Communication_PC".Para.DrillDepth - 5.0);

   // ---------- 网络 5 ----------
   // 标题：流程启动
   // 含义：将 ((((((((#DownDrillStep.StartCmd AND #DownDrillStep.OKToStart) OR #DownDrillStep.StepStart) AND "AllMode_M") AND "DB1900_Communication_PC".Recv.Z05ExtTPPB) AND ("DB1900_Communication_PC".Recv.Current_2 >= 0.5))) AND NOT ("DB1900_Communication_PC".Recv.EmmMode)) AND NOT ("DB1040_HomePos".Status.Running)) AND NOT (#DownDrillStep.StepEnd) 赋给 #DownDrillStep.StepStart
   #DownDrillStep.StepStart := ((((((((#DownDrillStep.StartCmd AND #DownDrillStep.OKToStart) OR #DownDrillStep.StepStart) AND "AllMode_M") AND "DB1900_Communication_PC".Recv.Z05ExtTPPB) AND ("DB1900_Communication_PC".Recv.Current_2 >= 0.5))) AND NOT ("DB1900_Communication_PC".Recv.EmmMode)) AND NOT ("DB1040_HomePos".Status.Running)) AND NOT (#DownDrillStep.StepEnd);
   // 含义：将 ((((((((#DownDrillStep.StartCmd AND #DownDrillStep.OKToStart) OR #DownDrillStep.StepStart) AND "AllMode_M") AND "DB1900_Communication_PC".Recv.Z05ExtTPPB) AND ("DB1900_Communication_PC".Recv.Current_2 >= 0.5))) AND NOT ("DB1900_Communication_PC".Recv.EmmMode)) AND NOT ("DB1040_HomePos".Status.Running)) AND NOT (#DownDrillStep.StepEnd) 赋给 #DownDrillStep.Busy
   #DownDrillStep.Busy := ((((((((#DownDrillStep.StartCmd AND #DownDrillStep.OKToStart) OR #DownDrillStep.StepStart) AND "AllMode_M") AND "DB1900_Communication_PC".Recv.Z05ExtTPPB) AND ("DB1900_Communication_PC".Recv.Current_2 >= 0.5))) AND NOT ("DB1900_Communication_PC".Recv.EmmMode)) AND NOT ("DB1040_HomePos".Status.Running)) AND NOT (#DownDrillStep.StepEnd);
   // 含义：条件 NOT (((((((((#DownDrillStep.StartCmd AND #DownDrillStep.OKToStart) OR #DownDrillStep.StepStart) AND "AllMode_M") AND "DB1900_Communication_PC".Recv.Z05ExtTPPB) AND ("DB1900_Communication_PC".Recv.Current_2 >= 0.5))) AND NOT ("DB1900_Communication_PC".Recv.EmmMode)) AND NOT ("DB1040_HomePos".Status.Running)) AND NOT (#DownDrillStep.StepEnd)) 成立时，将 FALSE 传送到 #DownDrillStep.ErrEnd
   IF NOT (((((((((#DownDrillStep.StartCmd AND #DownDrillStep.OKToStart) OR #DownDrillStep.StepStart) AND "AllMode_M") AND "DB1900_Communication_PC".Recv.Z05ExtTPPB) AND ("DB1900_Communication_PC".Recv.Current_2 >= 0.5))) AND NOT ("DB1900_Communication_PC".Recv.EmmMode)) AND NOT ("DB1040_HomePos".Status.Running)) AND NOT (#DownDrillStep.StepEnd)) THEN
       #DownDrillStep.ErrEnd := FALSE;
   END_IF;
   // 含义：条件 NOT (((((((((#DownDrillStep.StartCmd AND #DownDrillStep.OKToStart) OR #DownDrillStep.StepStart) AND "AllMode_M") AND "DB1900_Communication_PC".Recv.Z05ExtTPPB) AND ("DB1900_Communication_PC".Recv.Current_2 >= 0.5))) AND NOT ("DB1900_Communication_PC".Recv.EmmMode)) AND NOT ("DB1040_HomePos".Status.Running)) AND NOT (#DownDrillStep.StepEnd)) 成立时，将 FALSE 传送到 #DownDrillStep.ByPass
   IF NOT (((((((((#DownDrillStep.StartCmd AND #DownDrillStep.OKToStart) OR #DownDrillStep.StepStart) AND "AllMode_M") AND "DB1900_Communication_PC".Recv.Z05ExtTPPB) AND ("DB1900_Communication_PC".Recv.Current_2 >= 0.5))) AND NOT ("DB1900_Communication_PC".Recv.EmmMode)) AND NOT ("DB1040_HomePos".Status.Running)) AND NOT (#DownDrillStep.StepEnd)) THEN
       #DownDrillStep.ByPass := FALSE;
   END_IF;
   // 含义：条件 NOT (((((((((#DownDrillStep.StartCmd AND #DownDrillStep.OKToStart) OR #DownDrillStep.StepStart) AND "AllMode_M") AND "DB1900_Communication_PC".Recv.Z05ExtTPPB) AND ("DB1900_Communication_PC".Recv.Current_2 >= 0.5))) AND NOT ("DB1900_Communication_PC".Recv.EmmMode)) AND NOT ("DB1040_HomePos".Status.Running)) AND NOT (#DownDrillStep.StepEnd)) 成立时，将 FALSE 传送到 #DownDrillStep.StopDrill_Ack
   IF NOT (((((((((#DownDrillStep.StartCmd AND #DownDrillStep.OKToStart) OR #DownDrillStep.StepStart) AND "AllMode_M") AND "DB1900_Communication_PC".Recv.Z05ExtTPPB) AND ("DB1900_Communication_PC".Recv.Current_2 >= 0.5))) AND NOT ("DB1900_Communication_PC".Recv.EmmMode)) AND NOT ("DB1040_HomePos".Status.Running)) AND NOT (#DownDrillStep.StepEnd)) THEN
       #DownDrillStep.StopDrill_Ack := FALSE;
   END_IF;

   // ---------- 网络 6 ----------
   // 标题：向下凿击模式
   // 含义：将 "DB1900_Communication_PC".Para.DrillDirection3 AND "DB1900_Communication_PC".Para.ProduceMode3 赋给 "DB720_KuKa_MainCtrl".CmdOut.di_DownChiselMode
   "DB720_KuKa_MainCtrl".CmdOut.di_DownChiselMode := "DB1900_Communication_PC".Para.DrillDirection3 AND "DB1900_Communication_PC".Para.ProduceMode3;

   // ---------- 网络 7 ----------
   // 标题：初始化
   // 含义：条件 ((#DownDrillStep.StepStart AND NOT (#DownDrillStep.ErrEnd)) AND NOT (#DownDrillStep.ByPass)) AND NOT (#DownDrillStep.S1) 成立时，将 FALSE 传送到 #DownDrillStep.TaskIO
   IF ((#DownDrillStep.StepStart AND NOT (#DownDrillStep.ErrEnd)) AND NOT (#DownDrillStep.ByPass)) AND NOT (#DownDrillStep.S1) THEN
       #DownDrillStep.TaskIO := FALSE;
   END_IF;
   // 含义：条件 ((#DownDrillStep.StepStart AND NOT (#DownDrillStep.ErrEnd)) AND NOT (#DownDrillStep.ByPass)) AND NOT (#DownDrillStep.S1) 成立时，将 FALSE 传送到 #DownDrillStep.TaskNIO
   IF ((#DownDrillStep.StepStart AND NOT (#DownDrillStep.ErrEnd)) AND NOT (#DownDrillStep.ByPass)) AND NOT (#DownDrillStep.S1) THEN
       #DownDrillStep.TaskNIO := FALSE;
   END_IF;
   // 含义：条件 ((#DownDrillStep.StepStart AND NOT (#DownDrillStep.ErrEnd)) AND NOT (#DownDrillStep.ByPass)) AND NOT (#DownDrillStep.S1) 成立时，将 FALSE 传送到 "DB720_KuKa_MainCtrl".CmdOut.di_ChiselCylinderRet
   IF ((#DownDrillStep.StepStart AND NOT (#DownDrillStep.ErrEnd)) AND NOT (#DownDrillStep.ByPass)) AND NOT (#DownDrillStep.S1) THEN
       "DB720_KuKa_MainCtrl".CmdOut.di_ChiselCylinderRet := FALSE;
   END_IF;
   // 含义：条件 ((#DownDrillStep.StepStart AND NOT (#DownDrillStep.ErrEnd)) AND NOT (#DownDrillStep.ByPass)) AND NOT (#DownDrillStep.S1) 成立时，将 FALSE 传送到 "DB720_KuKa_MainCtrl".CmdOut.di_ChiselRobotRet
   IF ((#DownDrillStep.StepStart AND NOT (#DownDrillStep.ErrEnd)) AND NOT (#DownDrillStep.ByPass)) AND NOT (#DownDrillStep.S1) THEN
       "DB720_KuKa_MainCtrl".CmdOut.di_ChiselRobotRet := FALSE;
   END_IF;
   // 含义：条件 ((#DownDrillStep.StepStart AND NOT (#DownDrillStep.ErrEnd)) AND NOT (#DownDrillStep.ByPass)) AND NOT (#DownDrillStep.S1) 成立时，将 FALSE 传送到 #DownDrillStep.StopDrill_Ack
   IF ((#DownDrillStep.StepStart AND NOT (#DownDrillStep.ErrEnd)) AND NOT (#DownDrillStep.ByPass)) AND NOT (#DownDrillStep.S1) THEN
       #DownDrillStep.StopDrill_Ack := FALSE;
   END_IF;
   // 含义：条件 ((#DownDrillStep.StepStart AND NOT (#DownDrillStep.ErrEnd)) AND NOT (#DownDrillStep.ByPass)) AND NOT (#DownDrillStep.S1) 成立时，将 1 传送到 "DB720_KuKa_MainCtrl".Aux.ForceNum
   IF ((#DownDrillStep.StepStart AND NOT (#DownDrillStep.ErrEnd)) AND NOT (#DownDrillStep.ByPass)) AND NOT (#DownDrillStep.S1) THEN
       "DB720_KuKa_MainCtrl".Aux.ForceNum := 1;
   END_IF;
   // 含义：将 (#DownDrillStep.StepStart AND NOT (#DownDrillStep.ErrEnd)) AND NOT (#DownDrillStep.ByPass) 赋给 #DownDrillStep.S1
   #DownDrillStep.S1 := (#DownDrillStep.StepStart AND NOT (#DownDrillStep.ErrEnd)) AND NOT (#DownDrillStep.ByPass);

   // ---------- 网络 8 ----------
   // 标题：判断条件
   // 含义：将 (#DownDrillStep.S1 AND NOT ("DB1147_PromptStartNotPmt".Public.ChangeDownloadSlab)) OR (#DownDrillStep.S1 AND #DownDrillStep.S2) 赋给 #DownDrillStep.S2
   #DownDrillStep.S2 := (#DownDrillStep.S1 AND NOT ("DB1147_PromptStartNotPmt".Public.ChangeDownloadSlab)) OR (#DownDrillStep.S1 AND #DownDrillStep.S2);
   // 含义：条件 #DownDrillStep.S1 AND "DB1147_PromptStartNotPmt".Public.ChangeDownloadSlab 成立时，将 TRUE 传送到 #DownDrillStep.ErrEnd
   IF #DownDrillStep.S1 AND "DB1147_PromptStartNotPmt".Public.ChangeDownloadSlab THEN
       #DownDrillStep.ErrEnd := TRUE;
   END_IF;

   // ---------- 网络 9 ----------
   // 标题：电源夹具ID号错误，请检查夹具！
   // 含义：将 ((((#DownDrillStep.S2 AND ("DB1900_Communication_PC".Para.IOFixtureNo = "DB1080_Component".IOFixtureIID.TP_CurFixtureID))) AND ("DB1900_Communication_PC".Para.PowerFixtureNo = "DB1080_Component".PowerFixtureID.TP_CurFixtureID))) OR (#DownDrillStep.S2 AND #DownDrillStep.S5) 赋给 #DownDrillStep.S5
   #DownDrillStep.S5 := ((((#DownDrillStep.S2 AND ("DB1900_Communication_PC".Para.IOFixtureNo = "DB1080_Component".IOFixtureIID.TP_CurFixtureID))) AND ("DB1900_Communication_PC".Para.PowerFixtureNo = "DB1080_Component".PowerFixtureID.TP_CurFixtureID))) OR (#DownDrillStep.S2 AND #DownDrillStep.S5);

   // ---------- 网络 10 ----------
   // 标题：推力气缸
   // 含义：条件 #DownDrillStep.S5 AND NOT (#DownDrillStep.S7) 成立时，将 TRUE 传送到 "DB1081_ValveCall".ST01.Z01.ExtAuto
   IF #DownDrillStep.S5 AND NOT (#DownDrillStep.S7) THEN
       "DB1081_ValveCall".ST01.Z01.ExtAuto := TRUE;
   END_IF;
   // 含义：条件 #DownDrillStep.S5 AND NOT (#DownDrillStep.S7) 成立时，将 TRUE 传送到 "DB1081_ValveCall".ST01.Z02.VentValveAuto
   IF #DownDrillStep.S5 AND NOT (#DownDrillStep.S7) THEN
       "DB1081_ValveCall".ST01.Z02.VentValveAuto := TRUE;
   END_IF;
   // 含义：条件 #DownDrillStep.S5 AND NOT (#DownDrillStep.S7) 成立时，将 TRUE 传送到 "DB1081_ValveCall".ST01.Z05.ExtAuto
   IF #DownDrillStep.S5 AND NOT (#DownDrillStep.S7) THEN
       "DB1081_ValveCall".ST01.Z05.ExtAuto := TRUE;
   END_IF;
   // 含义：条件 #DownDrillStep.S5 AND NOT (#DownDrillStep.S7) 成立时，将 TRUE 传送到 "DB1081_ValveCall".ST01.Z06.RetAuto
   IF #DownDrillStep.S5 AND NOT (#DownDrillStep.S7) THEN
       "DB1081_ValveCall".ST01.Z06.RetAuto := TRUE;
   END_IF;
   // 含义：条件 (((#DownDrillStep.S5 AND NOT (#DownDrillStep.S7)) AND ("DB720_KuKa_MainCtrl".CmdOut.gi_ToolTypeNo = 13))) AND TRUE 成立时，将 TRUE 传送到 "QCamCoverExt"
   IF (((#DownDrillStep.S5 AND NOT (#DownDrillStep.S7)) AND ("DB720_KuKa_MainCtrl".CmdOut.gi_ToolTypeNo = 13))) AND TRUE THEN
       "QCamCoverExt" := TRUE;
   END_IF;
   // 含义：条件 (((#DownDrillStep.S5 AND NOT (#DownDrillStep.S7)) AND ("DB720_KuKa_MainCtrl".CmdOut.gi_ToolTypeNo = 13))) AND TRUE 成立时，将 FALSE 传送到 "QCamCoverRet"
   IF (((#DownDrillStep.S5 AND NOT (#DownDrillStep.S7)) AND ("DB720_KuKa_MainCtrl".CmdOut.gi_ToolTypeNo = 13))) AND TRUE THEN
       "QCamCoverRet" := FALSE;
   END_IF;
   // 含义：条件 #DownDrillStep.S5 AND NOT (#DownDrillStep.S7) 成立时，将 0.0 传送到 "DB1900_Communication_PC".Send.ScrLen
   IF #DownDrillStep.S5 AND NOT (#DownDrillStep.S7) THEN
       "DB1900_Communication_PC".Send.ScrLen := 0.0;
   END_IF;
   // 含义：条件 #DownDrillStep.S5 AND NOT (#DownDrillStep.S7) 成立时，将 0.45 传送到 "DB1080_Component".Aux.Pressure
   IF #DownDrillStep.S5 AND NOT (#DownDrillStep.S7) THEN
       "DB1080_Component".Aux.Pressure := 0.45;
   END_IF;
   // 含义：将 ((#DownDrillStep.S5 AND "DB1081_ValveCall".ST01.Z01.ExtPos) AND "DB1081_ValveCall".ST01.Z06.RetPos) OR (#DownDrillStep.S5 AND #DownDrillStep.S7) 赋给 #DownDrillStep.S7
   #DownDrillStep.S7 := ((#DownDrillStep.S5 AND "DB1081_ValveCall".ST01.Z01.ExtPos) AND "DB1081_ValveCall".ST01.Z06.RetPos) OR (#DownDrillStep.S5 AND #DownDrillStep.S7);

   // ---------- 网络 11 ----------
   // 标题：数据写入 X宽 Y长
   // 注释：PosNo is ToolNo, not HoleNo.
   // 含义：将 "DB1910_DrillData".DownDrill.gi_OffSetY; (* Convert → DInt *) END_IF 赋给 IF #DownDrillStep.S7 AND NOT (#DownDrillStep.S10) THEN "DB720_KuKa_MainCtrl".Aux.OffSetYMid
   IF #DownDrillStep.S7 AND NOT (#DownDrillStep.S10) THEN
       "DB720_KuKa_MainCtrl".Aux.OffSetYMid := "DB1910_DrillData".DownDrill.gi_OffSetY; (* Convert → DInt *)
   END_IF;
   // 含义：将 SWAP("DB720_KuKa_MainCtrl".Aux.OffSetYMid) 赋给 "DB720_KuKa_MainCtrl".CmdOut.gi_OffSetY
   "DB720_KuKa_MainCtrl".CmdOut.gi_OffSetY := SWAP("DB720_KuKa_MainCtrl".Aux.OffSetYMid);
   // 含义：将 "DB1910_DrillData".DownDrill.gi_OffsetX; (* Convert → DInt *) END_IF 赋给 IF #DownDrillStep.S7 AND NOT (#DownDrillStep.S10) THEN "DB720_KuKa_MainCtrl".Aux.OffSetZMid
   IF #DownDrillStep.S7 AND NOT (#DownDrillStep.S10) THEN
       "DB720_KuKa_MainCtrl".Aux.OffSetZMid := "DB1910_DrillData".DownDrill.gi_OffsetX; (* Convert → DInt *)
   END_IF;
   // 含义：将 SWAP("DB720_KuKa_MainCtrl".Aux.OffSetZMid) 赋给 "DB720_KuKa_MainCtrl".CmdOut.gi_OffSetX
   "DB720_KuKa_MainCtrl".CmdOut.gi_OffSetX := SWAP("DB720_KuKa_MainCtrl".Aux.OffSetZMid);
   // 含义：将 "DB1900_Communication_PC".Para.ScrLen; (* Convert → DInt *) END_IF 赋给 IF #DownDrillStep.S7 AND NOT (#DownDrillStep.S10) THEN "DB720_KuKa_MainCtrl".Aux.ScrLen_Mid0
   IF #DownDrillStep.S7 AND NOT (#DownDrillStep.S10) THEN
       "DB720_KuKa_MainCtrl".Aux.ScrLen_Mid0 := "DB1900_Communication_PC".Para.ScrLen; (* Convert → DInt *)
   END_IF;
   // 含义：将 SWAP("DB720_KuKa_MainCtrl".Aux.ScrLen_Mid0) 赋给 "DB720_KuKa_MainCtrl".CmdOut.gi_ScrewLength
   "DB720_KuKa_MainCtrl".CmdOut.gi_ScrewLength := SWAP("DB720_KuKa_MainCtrl".Aux.ScrLen_Mid0);
   // 含义：当 #DownDrillStep.S7 为 TRUE 时置位 #DownDrillStep.S10，否则复位（触点→线圈）
   IF #DownDrillStep.S7 THEN
       #DownDrillStep.S10 := TRUE;
   ELSE
       #DownDrillStep.S10 := FALSE;
   END_IF;

   // ---------- 网络 12 ----------
   // 注释：Add M29.0 to Acclerate DownChisel 2023.0302
   // 含义：将 (((#DownDrillStep.S10 AND "IZ02ExtPos") AND ("DB1080_Component".ClinyderPos.Ctrl_Out.Cur_Val_Out <= 1.0))) OR ((#DownDrillStep.S10 AND "DB1900_Communication_PC".Para.DrillDirection3) AND "DB1900_Communication_PC".Para.ProduceMode3) OR (#DownDrillStep.S10 AND #DownDrillStep.S12) 赋给 #DownDrillStep.S12
   #DownDrillStep.S12 := (((#DownDrillStep.S10 AND "IZ02ExtPos") AND ("DB1080_Component".ClinyderPos.Ctrl_Out.Cur_Val_Out <= 1.0))) OR ((#DownDrillStep.S10 AND "DB1900_Communication_PC".Para.DrillDirection3) AND "DB1900_Communication_PC".Para.ProduceMode3) OR (#DownDrillStep.S10 AND #DownDrillStep.S12);
   // 含义：条件 (((((#DownDrillStep.S10 AND "DB1900_Communication_PC".Para.DrillDirection3) AND "DB1900_Communication_PC".Para.ProduceMode3) AND "IZ02ExtPos") AND "DB1081_ValveCall".ST01.Z01.ExtPos) AND ("DB1080_Component".ClinyderPos.Ctrl_Out.Cur_Val_Out <= 1.0)) 成立时，将 TRUE 传送到 "DB720_KuKa_MainCtrl".CmdOut.di_PushCylOK_Sig
   IF (((((#DownDrillStep.S10 AND "DB1900_Communication_PC".Para.DrillDirection3) AND "DB1900_Communication_PC".Para.ProduceMode3) AND "IZ02ExtPos") AND "DB1081_ValveCall".ST01.Z01.ExtPos) AND ("DB1080_Component".ClinyderPos.Ctrl_Out.Cur_Val_Out <= 1.0)) THEN
       "DB720_KuKa_MainCtrl".CmdOut.di_PushCylOK_Sig := TRUE;
   END_IF;
   // 含义：条件 (((#DownDrillStep.S10 AND "DB1900_Communication_PC".Para.DrillDirection3) AND "DB1900_Communication_PC".Para.ProduceMode3) AND ("DB1080_Component".ClinyderPos.Ctrl_Out.Cur_Val_Out > 1.0)) 成立时，将 FALSE 传送到 "DB720_KuKa_MainCtrl".CmdOut.di_PushCylOK_Sig
   IF (((#DownDrillStep.S10 AND "DB1900_Communication_PC".Para.DrillDirection3) AND "DB1900_Communication_PC".Para.ProduceMode3) AND ("DB1080_Component".ClinyderPos.Ctrl_Out.Cur_Val_Out > 1.0)) THEN
       "DB720_KuKa_MainCtrl".CmdOut.di_PushCylOK_Sig := FALSE;
   END_IF;

   // ---------- 网络 13 ----------
   // 标题：调用机器人
   // 含义：条件 (#DownDrillStep.S12 AND NOT (#DownDrillStep.S15)) AND NOT ("DB720_KuKa_MainCtrl".CmdOut.di_DownChiselMode) 成立时，将 3 传送到 "DB1080_Component".Robot.CTRL_IN.ProgNo
   IF (#DownDrillStep.S12 AND NOT (#DownDrillStep.S15)) AND NOT ("DB720_KuKa_MainCtrl".CmdOut.di_DownChiselMode) THEN
       "DB1080_Component".Robot.CTRL_IN.ProgNo := 3;
   END_IF;
   // 含义：条件 (#DownDrillStep.S12 AND NOT (#DownDrillStep.S15)) AND "DB720_KuKa_MainCtrl".CmdOut.di_DownChiselMode 成立时，将 16 传送到 "DB1080_Component".Robot.CTRL_IN.ProgNo
   IF (#DownDrillStep.S12 AND NOT (#DownDrillStep.S15)) AND "DB720_KuKa_MainCtrl".CmdOut.di_DownChiselMode THEN
       "DB1080_Component".Robot.CTRL_IN.ProgNo := 16;
   END_IF;
   // 含义：将 #DownDrillStep.S12 AND NOT (#DownDrillStep.S15) 赋给 "DB1146_PromptFree".Public.do_DownDril_Act
   "DB1146_PromptFree".Public.do_DownDril_Act := #DownDrillStep.S12 AND NOT (#DownDrillStep.S15);
   // 含义：条件 #DownDrillStep.S12 AND NOT (#DownDrillStep.S15) 成立时，将 30 传送到 "DB1080_Component".Robot.CTRL_IN.RobotSpeed
   IF #DownDrillStep.S12 AND NOT (#DownDrillStep.S15) THEN
       "DB1080_Component".Robot.CTRL_IN.RobotSpeed := 30;
   END_IF;
   // 含义：条件 #DownDrillStep.S12 成立时，将 TRUE 传送到 "DB1080_Component".Robot.Cmd.Auto.ProgStart
   IF #DownDrillStep.S12 THEN
       "DB1080_Component".Robot.Cmd.Auto.ProgStart := TRUE;
   END_IF;
   // 含义：将 (((#DownDrillStep.S12 AND "DB1081_ValveCall".ST01.Z05.ExtPos) AND "DB1080_Component".Robot.Status.Busy) AND "DB720_KuKa_MainCtrl".StatusIn.do_DownDril_Pos) OR (#DownDrillStep.S12 AND #DownDrillStep.S15) 赋给 #DownDrillStep.S15
   #DownDrillStep.S15 := (((#DownDrillStep.S12 AND "DB1081_ValveCall".ST01.Z05.ExtPos) AND "DB1080_Component".Robot.Status.Busy) AND "DB720_KuKa_MainCtrl".StatusIn.do_DownDril_Pos) OR (#DownDrillStep.S12 AND #DownDrillStep.S15);

   // ---------- 网络 14 ----------
   // 标题：钻孔数据
   // 含义：条件 ((#DownDrillStep.S15 AND NOT (#DownDrillStep.S20)) AND ("DB1910_DrillData".DownDrill.PosNo = 0)) 成立时，将 "DB1910_DrillData".DownDrill.CurrentDrillLength 传送到 "DB1910_DrillData".DownDrill.AlreadyDrillLength
   IF ((#DownDrillStep.S15 AND NOT (#DownDrillStep.S20)) AND ("DB1910_DrillData".DownDrill.PosNo = 0)) THEN
       "DB1910_DrillData".DownDrill.AlreadyDrillLength := "DB1910_DrillData".DownDrill.CurrentDrillLength;
   END_IF;
   // 含义：条件 ((#DownDrillStep.S15 AND NOT (#DownDrillStep.S20)) AND ("DB1910_DrillData".DownDrill.PosNo >= 1)) 成立时，将 ("DB1910_DrillData".DownDrill.AlreadyDrillLength + "DB1910_DrillData".DownDrill.CurrentDrillLength) 传送到 "DB1910_DrillData".DownDrill.AlreadyDrillLength
   IF ((#DownDrillStep.S15 AND NOT (#DownDrillStep.S20)) AND ("DB1910_DrillData".DownDrill.PosNo >= 1)) THEN
       "DB1910_DrillData".DownDrill.AlreadyDrillLength := ("DB1910_DrillData".DownDrill.AlreadyDrillLength + "DB1910_DrillData".DownDrill.CurrentDrillLength);
   END_IF;
   // 含义：条件 #DownDrillStep.S15 AND NOT (#DownDrillStep.S20) 成立时，将 ("DB1910_DrillData".DownDrill.PosNo + 1) 传送到 "DB1910_DrillData".DownDrill.PosNo
   IF #DownDrillStep.S15 AND NOT (#DownDrillStep.S20) THEN
       "DB1910_DrillData".DownDrill.PosNo := ("DB1910_DrillData".DownDrill.PosNo + 1);
   END_IF;
   // 含义：当 #DownDrillStep.S15 为 TRUE 时置位 #DownDrillStep.S20，否则复位（触点→线圈）
   IF #DownDrillStep.S15 THEN
       #DownDrillStep.S20 := TRUE;
   ELSE
       #DownDrillStep.S20 := FALSE;
   END_IF;
   // 含义：将 #DownDrillStep.S15 AND NOT (#DownDrillStep.S22) 赋给 "DB720_KuKa_MainCtrl".CmdOut.di_DownDril_Ack
   "DB720_KuKa_MainCtrl".CmdOut.di_DownDril_Ack := #DownDrillStep.S15 AND NOT (#DownDrillStep.S22);
   // 含义：条件 #DownDrillStep.S15 AND "DB720_KuKa_MainCtrl".StatusIn.do_DownDrilApp_Pos 成立时，将 TRUE 传送到 "DB1081_ValveCall".ST01.Z01.ExtAuto
   IF #DownDrillStep.S15 AND "DB720_KuKa_MainCtrl".StatusIn.do_DownDrilApp_Pos THEN
       "DB1081_ValveCall".ST01.Z01.ExtAuto := TRUE;
   END_IF;
   // 含义：条件 #DownDrillStep.S15 AND "DB720_KuKa_MainCtrl".StatusIn.do_DownDrilApp_Pos 成立时，将 TRUE 传送到 "DB1081_ValveCall".ST01.Z02.RetAuto
   IF #DownDrillStep.S15 AND "DB720_KuKa_MainCtrl".StatusIn.do_DownDrilApp_Pos THEN
       "DB1081_ValveCall".ST01.Z02.RetAuto := TRUE;
   END_IF;
   // 含义：条件 #DownDrillStep.S15 AND "DB720_KuKa_MainCtrl".StatusIn.do_DownDrilApp_Pos 成立时，将 0.3 传送到 "DB1080_Component".Aux.Pressure
   IF #DownDrillStep.S15 AND "DB720_KuKa_MainCtrl".StatusIn.do_DownDrilApp_Pos THEN
       "DB1080_Component".Aux.Pressure := 0.3;
   END_IF;

   // ---------- 网络 15 ----------
   // 标题：速度分时
   // 含义：本网络为 StructuredText（SCL）原文重建，非 LAD 折叠
   IF #Aux.StartDrill AND
       NOT #DownDrillStep.S22 AND
       NOT "DB720_KuKa_MainCtrl".StatusIn.do_ReqStopDril AND
       "DB720_KuKa_MainCtrl".StatusIn.do_ReqDrilling
   THEN
       "DB720_KuKa_MainCtrl".Aux.RobotSpeed := REAL_TO_DINT("DB1080_Component".ClinyderPos.Ctrl_Out.Cur_Val_Out * (-1.0) + 100);
       IF "DB720_KuKa_MainCtrl".Aux.RobotSpeed > 35
       THEN
           "DB1080_Component".Robot.CTRL_IN.RobotSpeed := DINT_TO_BYTE(("DB720_KuKa_MainCtrl".Aux.RobotSpeed) * "DB1900_Communication_PC".Para.RobotSpeed / 100);
       ELSE
           "DB1080_Component".Robot.CTRL_IN.RobotSpeed := 30;
       END_IF;
   END_IF;
   IF "DB720_KuKa_MainCtrl".StatusIn.do_DownDril_Pos THEN
       IF "DB1900_Communication_PC".Para.CurrentMaxLimit > 5.0 THEN
           IF "DB1900_Communication_PC".Recv.Current_2 > ("DB1900_Communication_PC".Para.CurrentMaxLimit - 1.5) THEN
               "DB1080_Component".Robot.CTRL_IN.RobotSpeed := 5;
           END_IF;
       ELSE
           IF "DB1900_Communication_PC".Recv.Current_2 > ("DB1900_Communication_PC".Para.CurrentMaxLimit - 0.5) THEN
               "DB1080_Component".Robot.CTRL_IN.RobotSpeed := 5;
           END_IF;
       END_IF;
   END_IF;

   // ---------- 网络 16 ----------
   // 标题：深度计算
   // 含义：条件 ((((((#DownDrillStep.S12 AND "DB720_KuKa_MainCtrl".StatusIn.do_DrillReady_Act) AND ("DB1900_Communication_PC".Recv.Current_2 > "DB1900_Communication_PC".Para.CurrentMinLimit))) OR ((#DownDrillStep.S12 AND "DB720_KuKa_MainCtrl".StatusIn.do_DrillReady_Act) AND "DB720_KuKa_MainCtrl".StatusIn.do_DownDril_Pos)) AND NOT ("DB1900_Communication_PC".Para.ProduceMode3)) OR ((((((#DownDrillStep.S12 AND "DB720_KuKa_MainCtrl".StatusIn.do_DrillReady_Act) AND ("DB1900_Communication_PC".Recv.Current_2 > "DB1900_Communication_PC".Para.CurrentMinLimit))) OR ((#DownDrillStep.S12 AND "DB720_KuKa_MainCtrl".StatusIn.do_DrillReady_Act) AND "DB720_KuKa_MainCtrl".StatusIn.do_DownDril_Pos)) AND "DB1900_Communication_PC".Para.ProduceMode3) AND NOT ("DB720_KuKa_MainCtrl".StatusIn.do_ChiselPry)) OR ((#DownDrillStep.S12 AND NOT (#DownDrillStep.S22)) AND #Aux.StartDrill)) AND NOT (#Aux.StartDrill) 成立时，将 "DB720_KuKa_MainCtrl".Aux.go_Z 传送到 "DB720_KuKa_MainCtrl".Aux.XZeroPos
   IF ((((((#DownDrillStep.S12 AND "DB720_KuKa_MainCtrl".StatusIn.do_DrillReady_Act) AND ("DB1900_Communication_PC".Recv.Current_2 > "DB1900_Communication_PC".Para.CurrentMinLimit))) OR ((#DownDrillStep.S12 AND "DB720_KuKa_MainCtrl".StatusIn.do_DrillReady_Act) AND "DB720_KuKa_MainCtrl".StatusIn.do_DownDril_Pos)) AND NOT ("DB1900_Communication_PC".Para.ProduceMode3)) OR ((((((#DownDrillStep.S12 AND "DB720_KuKa_MainCtrl".StatusIn.do_DrillReady_Act) AND ("DB1900_Communication_PC".Recv.Current_2 > "DB1900_Communication_PC".Para.CurrentMinLimit))) OR ((#DownDrillStep.S12 AND "DB720_KuKa_MainCtrl".StatusIn.do_DrillReady_Act) AND "DB720_KuKa_MainCtrl".StatusIn.do_DownDril_Pos)) AND "DB1900_Communication_PC".Para.ProduceMode3) AND NOT ("DB720_KuKa_MainCtrl".StatusIn.do_ChiselPry)) OR ((#DownDrillStep.S12 AND NOT (#DownDrillStep.S22)) AND #Aux.StartDrill)) AND NOT (#Aux.StartDrill) THEN
       "DB720_KuKa_MainCtrl".Aux.XZeroPos := "DB720_KuKa_MainCtrl".Aux.go_Z;
   END_IF;
   // 含义：条件 (((((#DownDrillStep.S12 AND "DB720_KuKa_MainCtrl".StatusIn.do_DrillReady_Act) AND ("DB1900_Communication_PC".Recv.Current_2 > "DB1900_Communication_PC".Para.CurrentMinLimit))) OR ((#DownDrillStep.S12 AND "DB720_KuKa_MainCtrl".StatusIn.do_DrillReady_Act) AND "DB720_KuKa_MainCtrl".StatusIn.do_DownDril_Pos)) AND NOT ("DB1900_Communication_PC".Para.ProduceMode3)) OR ((((((#DownDrillStep.S12 AND "DB720_KuKa_MainCtrl".StatusIn.do_DrillReady_Act) AND ("DB1900_Communication_PC".Recv.Current_2 > "DB1900_Communication_PC".Para.CurrentMinLimit))) OR ((#DownDrillStep.S12 AND "DB720_KuKa_MainCtrl".StatusIn.do_DrillReady_Act) AND "DB720_KuKa_MainCtrl".StatusIn.do_DownDril_Pos)) AND "DB1900_Communication_PC".Para.ProduceMode3) AND NOT ("DB720_KuKa_MainCtrl".StatusIn.do_ChiselPry)) OR ((#DownDrillStep.S12 AND NOT (#DownDrillStep.S22)) AND #Aux.StartDrill) 成立时，将 ("DB720_KuKa_MainCtrl".Aux.go_Z - "DB720_KuKa_MainCtrl".Aux.XZeroPos) 传送到 "DB720_KuKa_MainCtrl".Aux.CurrentRobPos
   IF (((((#DownDrillStep.S12 AND "DB720_KuKa_MainCtrl".StatusIn.do_DrillReady_Act) AND ("DB1900_Communication_PC".Recv.Current_2 > "DB1900_Communication_PC".Para.CurrentMinLimit))) OR ((#DownDrillStep.S12 AND "DB720_KuKa_MainCtrl".StatusIn.do_DrillReady_Act) AND "DB720_KuKa_MainCtrl".StatusIn.do_DownDril_Pos)) AND NOT ("DB1900_Communication_PC".Para.ProduceMode3)) OR ((((((#DownDrillStep.S12 AND "DB720_KuKa_MainCtrl".StatusIn.do_DrillReady_Act) AND ("DB1900_Communication_PC".Recv.Current_2 > "DB1900_Communication_PC".Para.CurrentMinLimit))) OR ((#DownDrillStep.S12 AND "DB720_KuKa_MainCtrl".StatusIn.do_DrillReady_Act) AND "DB720_KuKa_MainCtrl".StatusIn.do_DownDril_Pos)) AND "DB1900_Communication_PC".Para.ProduceMode3) AND NOT ("DB720_KuKa_MainCtrl".StatusIn.do_ChiselPry)) OR ((#DownDrillStep.S12 AND NOT (#DownDrillStep.S22)) AND #Aux.StartDrill) THEN
       "DB720_KuKa_MainCtrl".Aux.CurrentRobPos := ("DB720_KuKa_MainCtrl".Aux.go_Z - "DB720_KuKa_MainCtrl".Aux.XZeroPos);
   END_IF;
   // 含义：将 ("DB720_KuKa_MainCtrl".Aux.CurrentRobPos - "DB1080_Component".ClinyderPos.Ctrl_Out.Cur_Val_Out) 赋给 "DB720_KuKa_MainCtrl".Aux.ScrLen_Mid1
   "DB720_KuKa_MainCtrl".Aux.ScrLen_Mid1 := ("DB720_KuKa_MainCtrl".Aux.CurrentRobPos - "DB1080_Component".ClinyderPos.Ctrl_Out.Cur_Val_Out);
   // 含义：条件 ("DB720_KuKa_MainCtrl".Aux.ScrLen_Mid1 >= 0.0) 成立时，将 "DB720_KuKa_MainCtrl".Aux.ScrLen_Mid1 传送到 "DB1900_Communication_PC".Send.ScrLen
   IF ("DB720_KuKa_MainCtrl".Aux.ScrLen_Mid1 >= 0.0) THEN
       "DB1900_Communication_PC".Send.ScrLen := "DB720_KuKa_MainCtrl".Aux.ScrLen_Mid1;
   END_IF;
   // 含义：将 (((((#DownDrillStep.S12 AND "DB720_KuKa_MainCtrl".StatusIn.do_DrillReady_Act) AND ("DB1900_Communication_PC".Recv.Current_2 > "DB1900_Communication_PC".Para.CurrentMinLimit))) OR ((#DownDrillStep.S12 AND "DB720_KuKa_MainCtrl".StatusIn.do_DrillReady_Act) AND "DB720_KuKa_MainCtrl".StatusIn.do_DownDril_Pos)) AND NOT ("DB1900_Communication_PC".Para.ProduceMode3)) OR ((((((#DownDrillStep.S12 AND "DB720_KuKa_MainCtrl".StatusIn.do_DrillReady_Act) AND ("DB1900_Communication_PC".Recv.Current_2 > "DB1900_Communication_PC".Para.CurrentMinLimit))) OR ((#DownDrillStep.S12 AND "DB720_KuKa_MainCtrl".StatusIn.do_DrillReady_Act) AND "DB720_KuKa_MainCtrl".StatusIn.do_DownDril_Pos)) AND "DB1900_Communication_PC".Para.ProduceMode3) AND NOT ("DB720_KuKa_MainCtrl".StatusIn.do_ChiselPry)) OR ((#DownDrillStep.S12 AND NOT (#DownDrillStep.S22)) AND #Aux.StartDrill) 赋给 #Aux.StartDrill
   #Aux.StartDrill := (((((#DownDrillStep.S12 AND "DB720_KuKa_MainCtrl".StatusIn.do_DrillReady_Act) AND ("DB1900_Communication_PC".Recv.Current_2 > "DB1900_Communication_PC".Para.CurrentMinLimit))) OR ((#DownDrillStep.S12 AND "DB720_KuKa_MainCtrl".StatusIn.do_DrillReady_Act) AND "DB720_KuKa_MainCtrl".StatusIn.do_DownDril_Pos)) AND NOT ("DB1900_Communication_PC".Para.ProduceMode3)) OR ((((((#DownDrillStep.S12 AND "DB720_KuKa_MainCtrl".StatusIn.do_DrillReady_Act) AND ("DB1900_Communication_PC".Recv.Current_2 > "DB1900_Communication_PC".Para.CurrentMinLimit))) OR ((#DownDrillStep.S12 AND "DB720_KuKa_MainCtrl".StatusIn.do_DrillReady_Act) AND "DB720_KuKa_MainCtrl".StatusIn.do_DownDril_Pos)) AND "DB1900_Communication_PC".Para.ProduceMode3) AND NOT ("DB720_KuKa_MainCtrl".StatusIn.do_ChiselPry)) OR ((#DownDrillStep.S12 AND NOT (#DownDrillStep.S22)) AND #Aux.StartDrill);
   // 含义：调用计数器实例 "DB1042_Timer".DDrillEndTime.TON（上升沿计数，当前值写入 CV）
   "DB1042_Timer".DDrillEndTime.TON(IN := (((((#DownDrillStep.S12 AND "DB720_KuKa_MainCtrl".StatusIn.do_DrillReady_Act) AND ("DB1900_Communication_PC".Recv.Current_2 > "DB1900_Communication_PC".Para.CurrentMinLimit))) OR ((#DownDrillStep.S12 AND "DB720_KuKa_MainCtrl".StatusIn.do_DrillReady_Act) AND "DB720_KuKa_MainCtrl".StatusIn.do_DownDril_Pos)) AND NOT ("DB1900_Communication_PC".Para.ProduceMode3)) OR ((((((#DownDrillStep.S12 AND "DB720_KuKa_MainCtrl".StatusIn.do_DrillReady_Act) AND ("DB1900_Communication_PC".Recv.Current_2 > "DB1900_Communication_PC".Para.CurrentMinLimit))) OR ((#DownDrillStep.S12 AND "DB720_KuKa_MainCtrl".StatusIn.do_DrillReady_Act) AND "DB720_KuKa_MainCtrl".StatusIn.do_DownDril_Pos)) AND "DB1900_Communication_PC".Para.ProduceMode3) AND NOT ("DB720_KuKa_MainCtrl".StatusIn.do_ChiselPry)) OR ((#DownDrillStep.S12 AND NOT (#DownDrillStep.S22)) AND #Aux.StartDrill),
                                    PT := "DB1900_Communication_PC".Para.DrillTime);

   // ---------- 网络 17 ----------
   // 标题：停止钻孔确认 后开始退枪 直到结束
   // 含义：条件 (((((#DownDrillStep.S20 AND NOT (#DownDrillStep.S22)) AND "DB720_KuKa_MainCtrl".StatusIn.do_ReqStopDril) AND ("DB1900_Communication_PC".Send.ScrLen > #Aux.DrillDepthMin))) AND NOT ("DB1900_Communication_PC".Para.DrillEndMode)) OR ((((#DownDrillStep.S20 AND NOT (#DownDrillStep.S22)) AND "DB720_KuKa_MainCtrl".StatusIn.do_ReqStopDril) AND "DB1042_Timer".DDrillEndTime.Q) AND "DB1900_Communication_PC".Para.DrillEndMode) OR ((#DownDrillStep.S20 AND NOT (#DownDrillStep.S22)) AND #DownDrillStep.StopDrill_End) 成立时，将 TRUE 传送到 #DownDrillStep.StopDrill_Ack
   IF (((((#DownDrillStep.S20 AND NOT (#DownDrillStep.S22)) AND "DB720_KuKa_MainCtrl".StatusIn.do_ReqStopDril) AND ("DB1900_Communication_PC".Send.ScrLen > #Aux.DrillDepthMin))) AND NOT ("DB1900_Communication_PC".Para.DrillEndMode)) OR ((((#DownDrillStep.S20 AND NOT (#DownDrillStep.S22)) AND "DB720_KuKa_MainCtrl".StatusIn.do_ReqStopDril) AND "DB1042_Timer".DDrillEndTime.Q) AND "DB1900_Communication_PC".Para.DrillEndMode) OR ((#DownDrillStep.S20 AND NOT (#DownDrillStep.S22)) AND #DownDrillStep.StopDrill_End) THEN
       #DownDrillStep.StopDrill_Ack := TRUE;
   END_IF;
   // 含义：将 ((#DownDrillStep.S20 AND NOT ("DB1900_Communication_PC".Para.ProduceMode3)) AND "DB720_KuKa_MainCtrl".StatusIn.do_DownDril_Don) OR ((#DownDrillStep.S20 AND "DB1900_Communication_PC".Para.ProduceMode3) AND "DB720_KuKa_MainCtrl".StatusIn.do_Gouge_Don) OR ((#DownDrillStep.S20 AND "DB1900_Communication_PC".Para.ProduceMode3) AND "DB720_KuKa_MainCtrl".StatusIn.do_Gouge_Don1) OR ((#DownDrillStep.S20 AND "DB1900_Communication_PC".Para.ProduceMode3) AND "DB720_KuKa_MainCtrl".StatusIn.do_DownDril_Don) OR (#DownDrillStep.S20 AND #DownDrillStep.S22) 赋给 #DownDrillStep.S22
   #DownDrillStep.S22 := ((#DownDrillStep.S20 AND NOT ("DB1900_Communication_PC".Para.ProduceMode3)) AND "DB720_KuKa_MainCtrl".StatusIn.do_DownDril_Don) OR ((#DownDrillStep.S20 AND "DB1900_Communication_PC".Para.ProduceMode3) AND "DB720_KuKa_MainCtrl".StatusIn.do_Gouge_Don) OR ((#DownDrillStep.S20 AND "DB1900_Communication_PC".Para.ProduceMode3) AND "DB720_KuKa_MainCtrl".StatusIn.do_Gouge_Don1) OR ((#DownDrillStep.S20 AND "DB1900_Communication_PC".Para.ProduceMode3) AND "DB720_KuKa_MainCtrl".StatusIn.do_DownDril_Don) OR (#DownDrillStep.S20 AND #DownDrillStep.S22);
   // 含义：条件 ((#DownDrillStep.S20 AND NOT ("DB1900_Communication_PC".Para.ProduceMode3)) AND "DB720_KuKa_MainCtrl".StatusIn.do_DownDril_Don) OR ((#DownDrillStep.S20 AND "DB1900_Communication_PC".Para.ProduceMode3) AND "DB720_KuKa_MainCtrl".StatusIn.do_Gouge_Don) OR ((#DownDrillStep.S20 AND "DB1900_Communication_PC".Para.ProduceMode3) AND "DB720_KuKa_MainCtrl".StatusIn.do_Gouge_Don1) OR ((#DownDrillStep.S20 AND "DB1900_Communication_PC".Para.ProduceMode3) AND "DB720_KuKa_MainCtrl".StatusIn.do_DownDril_Don) OR (#DownDrillStep.S20 AND #DownDrillStep.S22) 成立时，将 FALSE 传送到 #DownDrillStep.StopDrill_Ack
   IF ((#DownDrillStep.S20 AND NOT ("DB1900_Communication_PC".Para.ProduceMode3)) AND "DB720_KuKa_MainCtrl".StatusIn.do_DownDril_Don) OR ((#DownDrillStep.S20 AND "DB1900_Communication_PC".Para.ProduceMode3) AND "DB720_KuKa_MainCtrl".StatusIn.do_Gouge_Don) OR ((#DownDrillStep.S20 AND "DB1900_Communication_PC".Para.ProduceMode3) AND "DB720_KuKa_MainCtrl".StatusIn.do_Gouge_Don1) OR ((#DownDrillStep.S20 AND "DB1900_Communication_PC".Para.ProduceMode3) AND "DB720_KuKa_MainCtrl".StatusIn.do_DownDril_Don) OR (#DownDrillStep.S20 AND #DownDrillStep.S22) THEN
       #DownDrillStep.StopDrill_Ack := FALSE;
   END_IF;

